(* Counting distance *)
IF bCount
    AND NOT fbFileHandler.bFileRead
THEN
	lrNoRetainDistance := lrNoRetainDistance + lrDistance;
	stRetainDistance.lrAllOverDistance := stCacheRetainDistance.lrAllOverDistance + lrNoRetainDistance;
	stRetainDistance.lrAfterResetDistance := stCacheRetainDistance.lrAfterResetDistance + lrNoRetainDistance;
END_IF


(* Write / read  file *)
fbFileHandler(
	bEnable := TRUE,
	dwDataBuffer := ADR(stRetainDistance),
	udnDataBufLen := SIZEOF(stRetainDistance),
	tTimeout := tTimeout,
	bError => bError,
	udnErrNo => udnErrNo
);

rtReset(
	CLK := NOT bSave AND bReset
);
IF rtReset.Q
THEN
	stRetainDistance.lrAfterResetDistance := 0;
	lrNoRetainDistance := 0;
END_IF

rtDeleteAll(
	CLK := NOT bSave AND bDeleteAll
);
IF rtDeleteAll.Q
THEN
	stRetainDistance.lrAllOverDistance := 0;
	stRetainDistance.lrAfterResetDistance := 0;
	stCacheRetainDistance.lrAllOverDistance := 0;
	stCacheRetainDistance.lrAfterResetDistance := 0;
	lrNoRetainDistance := 0;
END_IF

(* Counter distance mapping *)
lrAllOverDistance := stRetainDistance.lrAllOverDistance;
lrAfterResetDistance := stRetainDistance.lrAfterResetDistance;

END_FUNCTION_BLOCK

// ---- POUs/Tc2 Objects/Measurements/FB_TemperaturOK.TcPOU
FUNCTION_BLOCK FB_TemperaturOK
VAR_INPUT
	bEnable						:BOOL;			(* Enable FB signal *)
	bIn							:BOOL;			(* Temperature OK *)
	tTimeOutTempOK				:TIME := t#5s;		(* Temperature OK timeout *)
	tTimeOutTempNOK			:TIME := t#5s;		(* Temperature NOK timeout *)
END_VAR
VAR_OUTPUT
	bOut					:BOOL;			(* Temperature OK *)
	bError					:BOOL;			(* Error by temperature NOK *)
	udnErrorNo				:UDINT;
	udnMessageNo			:UDINT;
	sMsg					:STRING;
END_VAR
VAR
	bFirstTime			:BOOL;			(* First cycle *)
	tonDelayOK			:TON;			(* Temperatur delay ok *)
	tofWatchDog			:TOF;			(* Timer to off *)

END_VAR


IF NOT bFirstTime
THEN
	bError := FALSE;
	udnErrorNo := 0;
	udnMessageNo := 0;
	sMsg := '';
	tonDelayOK(
		IN := FALSE,
	          PT := tTimeOutTempOK
	);
	tofWatchDog(
		IN := FALSE,
	         PT := tTimeOutTempNOK
	);
	bFirstTime := TRUE;
END_IF;

(* Timer starts when came rising edge of signal *)
tonDelayOK(
	IN := bIn,
         PT := tTimeOutTempOK
);

tofWatchDog(
	IN := bIn,
         PT := tTimeOutTempNOK
);

IF tonDelayOK.Q
THEN
	bOut := TRUE;
    
ELSIF NOT tofWatchDog.Q
THEN
	bOut := FALSE;
    
END_IF;

END_FUNCTION_BLOCK

// ---- POUs/Tc2 Objects/Measurements/Oscat/T_PLC_MS.TcPOU
FUNCTION T_PLC_MS : DWORD
VAR CONSTANT
	debug			:BOOL := 0;
	N 				:INT := 0;
	offset 			:DWORD := 0;
END_VAR
VAR
	tx 				:TIME;
END_VAR

(*
version 1.2	16. nov 2008
programmer 	hugo
tested by	oscat

T_PLC_MS reads the internal PLC timer and return the time, it has the advantage to be able to set a debug mode 
and speed up the counter to test the plc timer overrun which occurs every 50 days respectively 25 days at siemens S7
this routine also allows to correct the behavior of s7 where the internal plc counter will not count all 32 bits.

*)

tx := TIME();
T_PLC_MS := TIME_TO_DWORD(Tx);
(* hier muss die korrektur für step7 stattfinden
plctime muss den vollen wertebereich von time ausnutzen:
wenn bei step7 time -24tage bis plus 24 tage ist dann muss der timer auch beim überlauf auf -24tage springen 
und auf keinen fall auf 0 !!!!
für siemens muss ein weiterer fb im main eingebunden werden der sicherstellt das alle 32 bits durchgezählt werden.
es kann nur ein fb sein den er muss sich das oberste (32te) bit merken.
oder etwa spring s7 bei überlauf auf -24 tage????? dann wäre keine korrektur nötig.
*)
IF debug
THEN
	T_PLC_MS := (SHL(T_PLC_MS,N) OR SHL(DWORD#1,N)-1) + OFFSET;
END_IF;

END_FUNCTION

// ---- POUs/Tc2 Objects/Safety/Fieldbus/FB_Fieldbus.TcPOU
FUNCTION_BLOCK FB_Fieldbus
(*

The function block used to control fieldbus.

Constructor: 		Patryk Panylo
Company:		E. Riexinger GmbH
Date:			23.04.2015
Version:			1.00

Date:			Revision:		Who:				Comment
dd.mm.yyyy		x.xx			Initials			comment

*)
VAR_INPUT
	(* Input variables / Eingang Variablen *)
	bEnable					:BOOL;						(* Enable FB signal *)
	unMasterState			:UINT;						(* Master state of fieldbus *)
														(* unFieldbus = 1 -> Sercos-Master:
															0xE001 = Phase 0
															0xE002 = Phase 1
															0xE003 = Phase 2
															0xE004 = Phase 3
															0xE005 = Phase 4
															0xE008 = Break
															0xE011 = Phase switch 0 -> 1
															0xE012 = Phase switch 1 -> 2
															0xE013 = Phase switch 2 -> 3
															0xE014 = Phase switch 3 -> 4
					
														  uiFieldbus = 2 -> EtherCat Master:
															0x0001 = Link error
															0x0002 = I/O locked after link error (I/O reset required)
															0x0004 = Link error (redundancy adapter)
															0x0008 = Missing one frame (redundancy mode)
															0x0010 = Out of send resources (I/O reset required)
															0x0020 = Watchdog triggered
															0x0040 = Ethernet driver (miniport) not found
															0x0080 = I/O reset active
															0x0100 = At least one device in 'INIT' state
															0x0200 = At least one device in 'PRE-OP' state
															0x0400 = At least one device in 'SAFE-OP' state
															0x0800 = At least one device indicates an error state
															0x1000 = DC not in sync
														*)
	unSlaveState				:ARRAY[1..unSlaveNo] OF UINT;	(* State of slaves periphery / Status des Periphery
														uiFieldbus = 2 -> EtherCat Master:
															0x___1 = Slave in 'INIT' state
															0x___2 = Slave in 'PREOP' state
															0x___3 = Slave in 'BOOT' state
															0x___4 = Slave in 'SAFEOP' state
															0x___8 = Slave in 'OP' state
															0x001_ = Slave signals error
															0x002_ = Invalid vendorId, productCode... read
															0x004_ = Initialization error occurred
															0x008_ = Slave disabled
															0x010_ = Slave not present
															0x020_ = Slave signals link error
															0x040_ = Slave signals missing link
															0x080_ = Slave signals unexpected link
															0x100_ = Communication port A
															0x200_ = Communication port B
															0x400_ = Communication port C
															0x800_ = Communication port D
													*)
	tAdsTimeOut				:TIME := t#5s;				(* Timeout for ADS commando *)
END_VAR
VAR_OUTPUT
	(* Output variables / Ausgang Variablen *)
	sDeviceNetId				:T_AmsNetId ;			(* Fieldbus master ams net id*)
	bInitReady				:BOOL;					(* Fieldbus master initialisation is complete*)
	bBreak					:BOOL;					(* Fieldbus break *)
	bError					:BOOL;					(* Error by no air pressure *)
	udnErrorNo				:UDINT;
	udnMessageNo			:UDINT;
	sMsg					:STRING;
END_VAR
VAR
	(* Enummerations *)

	(* Variables *)
	unSlaveCounter			:UINT;					(* Slave counter *)
	bBreakMasterState		:BOOL;					(* Fieldbus master break *)
	bBreakSlaveState			:BOOL;					(* Fieldbus slave break *)

	(* References *)

	(* Interfaces *)

	(* Instances *)
	fbGetDeviceNetId			:IOF_GetDeviceNetId; 		(* Get the device net id from the device ID *)
	fbGetDeviceType			:IOF_GetDeviceType; 		(* Get the device type from the device ID *)
END_VAR
VAR CONSTANT
	unSlaveNo				:UINT := 32;				(* Number of slaves in Fieldbus *)
END_VAR

IF NOT bEnable
THEN
	fbGetDeviceNetId(START := FALSE);
	fbGetDeviceType(START := FALSE);
	bInitReady := FALSE;
	bBreak := FALSE;
	bError := FALSE;
	udnErrorNo := 0;
	udnMessageNo := 0;
	sMsg := '';
	RETURN;
END_IF;

(* Get the device net id from the device ID *)
fbGetDeviceNetId(
	NETID := '',
	DEVICEID := 1,
	START := TRUE,
	TMOUT := tAdsTimeOut
);

(* Get the device type from the device ID *)
fbGetDeviceType(
	NETID := '',
	DEVICEID := 1,
	START := TRUE,
	TMOUT := tAdsTimeOut
);

(* Get the device net id from the device ID *)
IF NOT fbGetDeviceNetId.BUSY 											(* No error *)
     AND NOT fbGetDeviceNetId.ERR
THEN
	sDeviceNetId := fbGetDeviceNetId.DeviceNetId;							(* Device net id *)

	(* Get the device type from the device ID *)
	IF NOT fbGetDeviceType.BUSY 										(* No error *)
	     AND NOT fbGetDeviceType.ERR
	THEN

		CASE fbGetDeviceType.IODeviceType
		OF
			48: (* IODEVICETYPE_FC7500 	:= 48,  Beckhoff-SERCOS-PCI *)
				bError := FALSE;
				udnErrorNo := 0;											(* Error number *)
				bInitReady := unMasterState = 16#E005; 						(* Actual Phase is 4 *)
				bBreak := unMasterState = 16#E008;							(* Interrupt / Broke *)
			94: (* IODEVICETYPE_EtherCAT := 94,  Beckhoff-EtherCAT-PCI *)
				bError := FALSE;
				udnErrorNo := 0;											(* Error number *)
				bInitReady := unMasterState = 16#0000; 						(* Actual master state is OP *)

				bBreakMasterState :=  unMasterState <> 16#0000;				(* Fieldbus master break *)

				IF bInitReady
				THEN
					bBreakSlaveState := FALSE;							(* Fieldbus slave break *)

					FOR unSlaveCounter :=1 TO unSlaveNo
					DO
						bBreakSlaveState := unSlaveState[unSlaveCounter] <> 16#0000
										     AND unSlaveState[unSlaveCounter] <> 16#0008;

						IF bBreakSlaveState
						THEN
							EXIT;
						END_IF

					END_FOR;
				END_IF

				bBreak := bBreakMasterState 								(* Interrupt / Broke *)
						 OR bBreakSlaveState;

		ELSE (* IDLE *)
			bInitReady := FALSE;
			bBreak := FALSE;
			bError := TRUE;
			udnErrorNo := 1;																			(* Error number *)
			sMsg := CONCAT('Unidentified fieldbus:', DINT_TO_STRING(fbGetDeviceType.IODeviceType));		(* Description error *)
		END_CASE;

	ELSIF NOT fbGetDeviceType.BUSY
		   AND fbGetDeviceType.ERR
	THEN
		bError := TRUE;
		udnErrorNo := 2;																				(* Error number *)
		sMsg := CONCAT('Fehler beim Lesen über ADS: ', UDINT_TO_STRING(fbGetDeviceType.ERRID));		(* Description error *)
		fbGetDeviceType(START := FALSE);
	END_IF;

ELSIF NOT fbGetDeviceNetId.BUSY
	    AND fbGetDeviceNetId.ERR
THEN
	bError := TRUE;
	udnErrorNo := 3;																					(* Error number *)
	sMsg := CONCAT('Fehler beim Lesen über ADS: ', UDINT_TO_STRING(fbGetDeviceNetId.ERRID));			(* Description error *)
	fbGetDeviceNetId(START := FALSE);
END_IF;

END_FUNCTION_BLOCK

// ---- POUs/Tc2 Objects/Signals/Force Input/FB_ForceBit.TcPOU
FUNCTION_BLOCK FB_ForceBit
(*

Forcing the input bit through pointer.
IO variables in VAR_CONFIG are generated automatically by TwinCAT - read only
Matching variable must be with  %I* declarated.

Constructor: 		Patryk Panylo
Company:		E. Riexinger GmbH
Date:			28.10.2013
Version:			1.00

Date:			Revision:		Who:				Comment
dd.mm.yyyy		x.xx			Initials			comment

*)
VAR_INPUT
	bEnable						:BOOL; 							(* Enable FB *)
	dwBitAddr					:DWORD;						(* The address of input argument in a DWORD: BITADR(Input) where e.g Input = %IX0.1 *)
	bForceInState				:BOOL;							(* Force input state *)
	tDelayOn					:TIME;							(* Delay signal on *)
	tDelayOff						:TIME;							(* Delay signal off *)
END_VAR
VAR_OUTPUT
END_VAR
VAR
	pByteAddr					:POINTER TO BYTE;
	byCurrentInState				:BYTE;							(* Current input state *)
	byBitMask					:BYTE;

	tonDelayOn					:TON;
	tonDelayOff					:TOF;

END_VAR

IF NOT bEnable
THEN
	RETURN;
END_IF

(* Delay on signal *)
tonDelayOn(
	IN := bForceInState,
	PT := tDelayOn
);

(* Delay off signal *)
tonDelayOff(
	IN := tonDelayOn.Q,
	PT := tDelayOff
);

pByteAddr := ADR(%IB0) + (dwBitAddr / 8);
byCurrentInState := pByteAddr^;

byBitMask := SHL(BYTE#1, (dwBitAddr AND 2#00000111));

IF tonDelayOff.Q
THEN
	pByteAddr^ := byCurrentInState OR byBitMask;
ELSE
	pByteAddr^ := byCurrentInState AND NOT byBitMask;
END_IF

END_FUNCTION_BLOCK

// ---- POUs/Tc2 Objects/Signals/Force Input/FB_ForceByte.TcPOU
FUNCTION_BLOCK FB_ForceByte
(*

Forcing the input bit through pointer.
IO variables in VAR_CONFIG are generated automatically by TwinCAT - read only
Matching variable must be with  %I* declarated.

Constructor: 		Patryk Panylo
Company:		E. Riexinger GmbH
Date:			28.10.2013
Version:			1.00

Date:			Revision:		Who:				Comment
dd.mm.yyyy		x.xx			Initials			comment

*)
VAR_INPUT
	bEnable						:BOOL; 							(* Enable FB *)
	dwAddr						:DWORD;						(* The address of input argument in a DWORD: ADR(Input) where e.g Input = %IB *)
	bForceInState				:BOOL;							(* Force input state *)
	tDelayOn					:TIME;							(* Delay signal on *)
	tDelayOff						:TIME;							(* Delay signal off *)
END_VAR
VAR_OUTPUT
END_VAR
VAR
	pByteAddr					:POINTER TO BYTE;
	byCurrentInState				:BYTE;							(* Current input state *)
	byBitMask					:BYTE;

	tonDelayOn					:TON;
	tonDelayOff					:TOF;

END_VAR

IF NOT bEnable
THEN
	RETURN;
END_IF

(* Delay on signal *)
tonDelayOn(
	IN := bForceInState,
	PT := tDelayOn
);

(* Delay off signal *)
tonDelayOff(
	IN := tonDelayOn.Q,
	PT := tDelayOff
);

pByteAddr := dwAddr;
byCurrentInState := pByteAddr^;

byBitMask := 2#00000001;

IF tonDelayOff.Q
THEN
	pByteAddr^ := byCurrentInState OR byBitMask;
ELSE
	pByteAddr^ := byCurrentInState AND NOT byBitMask;
END_IF

END_FUNCTION_BLOCK

// ---- POUs/Tc2 Objects/Signals/Handling/F_SignalHandling.TcPOU
FUNCTION F_SignalHandling : BOOL
VAR_INPUT
	(* Input variables / Eingang Variablen *)
	bEnable					:BOOL;						(* Enable FB signal *)
	bIn						:BOOL;						(* Input signal *)
END_VAR
VAR
END_VAR

IF NOT bEnable
THEN
	F_SignalHandling := FALSE;
    	RETURN;
END_IF;

F_SignalHandling := bIn;                     (* Set output *)

END_FUNCTION

// ---- POUs/Tc2 Objects/Signals/Ramp Generators/FB_RampDirector.TcPOU
FUNCTION_BLOCK FB_RampDirector
(*

Frequency division

Constructor: 		Patryk Panylo
Company:		E. Riexinger GmbH
Date:			14.11.2012
Version:			1.00

Date:			Revision:		Who:				Comment
dd.mm.yyyy		x.xx			Initials			comment

*)

VAR_INPUT
	bEnable						:BOOL;						(* Function block enable *)
	bExecute					:BOOL;						(* Execut the function block *)
	bDirection					:BOOL;						(* Rising = 1, Falling = 0 *)
	bSet						:BOOL;						(* Set output to 65535 *)
	bReset						:BOOL;						(* Reset output to 0 *)
	tRiseTime					:TIME;						(* Rise time of ramp *)
	tFallTime					:TIME;						(* Fall time of ramp *)
	rHighLimit					:REAL;						(* High limit of ramp *)
	rLowLimit						:REAL;						(* Low limit of ramp *)
	rNoLimit						:REAL;						(* No limit value active if rise and fall time no active *)
END_VAR
VAR_OUTPUT
	wRVOut						:WORD;						(* Ramp value, 100% = 65535 *)
	rPVOut						:REAL;						(* Judgment Value *)
	nPVOut						:INT;						(* Judgment Value *)
	bLowLevel					:BOOL;						(* Low level reached *)
	bHighLevel					:BOOL;						(* High level reached *)
	bDone						:BOOL;						(* Program done *)
	bBusy 						:BOOL;						(* Program busy *)
	bError 						:BOOL;						(* Program error *)
END_VAR
VAR
	fbRampGen					:FB_RMP_W;					(* Ramp generator *)

	rCacheLowLimit				:REAL;
	rCacheHighLimit				:REAL;

	rtExecute						:R_TRIG;
	etRampGenerator				:ET_RampGenerator;
END_VAR


IF NOT bEnable
THEN
	bDone := FALSE;                                     (* Program done *)
	bBusy := FALSE;                                     (* Program not busy *)
	bError := FALSE;                                    (* Program not error *)
	
	rtExecute(CLK := FALSE);

	fbRampGen(
		bEnable := FALSE,
		bReset := bReset,
		bSet := bSet,
		wRVOut => wRVOut
	);

	RETURN;
END_IF;

rtExecute(CLK := bExecute);

IF rtExecute.Q
THEN
	fbRampGen(
		bEnable := FALSE,
		bDirection := bDirection,
		bSet := FALSE,
		bReset := FALSE,
		tRampTime := T#0ms
	);
	
	etRampGenerator := ET_RampGenerator_eWaitExecute;						(* Next step *)

END_IF

(* Reset ramp *)
IF (tFallTime = t#0s
    AND tRiseTime <> t#0s
    AND bExecute
    AND NOT bDirection)
    OR bReset
THEN
	fbRampGen.bReset := TRUE;
	wRVOut := fbRampGen.wRVOut;
ELSE
	fbRampGen.bReset := FALSE;
END_IF;

(* Set ramp *)
IF (tRiseTime = t#0s
    AND tFallTime <> t#0s
    AND bExecute
    AND bDirection)
    OR bSet
THEN
	fbRampGen.bSet := TRUE;
ELSE
	fbRampGen.bSet := FALSE;
END_IF;

(* Call ramp generator *)
fbRampGen(
	bDirection := bDirection,
	tRampTime := SEL(bDirection, tFallTime, tRiseTime),
	bLowLevel => bLowLevel,
	bHighLevel => bHighLevel
);

IF fbRampGen.bReset
    OR fbRampGen.bSet
THEN
	wRVOut := fbRampGen.wRVOut;
END_IF;

CASE etRampGenerator OF
        
	ET_RampGenerator_eWaitExecute:
		bDone := FALSE;                                     (* Program done *)
		bBusy := FALSE;                                     (* Program not  busy *)
		bError := FALSE;                                    (* Program not error *)

		fbRampGen.bEnable := FALSE;
		
		IF rtExecute.Q
		THEN
			bDone := FALSE;                                     (* Program done *)
			bBusy := TRUE;                                 	 	(* Program not busy *)

			IF tRiseTime = t#0s
    			     AND tFallTime = t#0s
			THEN
				fbRampGen.bEnable := FALSE;

				rCacheLowLimit := rNoLimit;
				rCacheHighLimit := rNoLimit;

				etRampGenerator := ET_RampGenerator_eDone;         (* Next step *)
			ELSE
				fbRampGen.bEnable := TRUE;

				rCacheLowLimit := rLowLimit;
				rCacheHighLimit := rHighLimit;

				etRampGenerator := ET_RampGenerator_eRunning;           (* Next step *)
			END_IF
		END_IF

	ET_RampGenerator_eRunning:
		IF fbRampGen.bBusy
		THEN
			wRVOut := fbRampGen.wRVOut;
		
			etRampGenerator := ET_RampGenerator_eWaiting;           (* Next step *)
		END_IF
        
	ET_RampGenerator_eWaiting:
		IF fbRampGen.bBusy
		THEN
			wRVOut := fbRampGen.wRVOut;
		ELSE
			fbRampGen.bEnable := FALSE;
		
			etRampGenerator := ET_RampGenerator_eDone;         (* Next step *)
		END_IF		

	ET_RampGenerator_eDone:
		bDone := TRUE;                                      (* Program done *)
		bBusy := FALSE;                                     (* Program not busy *)
		
		etRampGenerator := ET_RampGenerator_eNotExecute;            (* Next step *)
        
	ET_RampGenerator_eError:
		bDone := FALSE;                                     (* Program done *)
		bBusy := FALSE;                                     (* Program not busy *)
		bError := TRUE;                                     (* Program error *)
		
		etRampGenerator := ET_RampGenerator_eNotExecute;            (* Next step *)
        
	ET_RampGenerator_eNotExecute:
	IF NOT bExecute
	THEN
		bDone := FALSE;                                     (* Program done *)
		bBusy := FALSE;                                     (* Program not busy *)
		bError := FALSE;                                    (* Program not error *)

		wRVOut := fbRampGen.wRVOut;
	
		etRampGenerator := ET_RampGenerator_eWaitExecute;               (* Next step *)

	END_IF;
END_CASE;

rPVOut := F_WordToRange(
			wWord := wRVOut,
			rLowLimit := rCacheLowLimit,
			rHighLimit := rCacheHighLimit
		);

nPVOut := REAL_TO_INT(rPVOut);

END_FUNCTION_BLOCK

// ---- POUs/Tc2 Objects/Signals/Watchdog/FB_SignalWatchdog2.TcPOU
FUNCTION_BLOCK FB_SignalWatchdog2
VAR_INPUT
	bEnable					:BOOL;			(* Enable FB signal *)
	bIn						:BOOL;			(* Input *)
	tTimeOutHigh				:TIME := t#5s;		(* Input high timeout *)
	tTimeOutLow				:TIME := t#5s;		(* Input low timeout *)
END_VAR
VAR_OUTPUT
	bOut					:BOOL;			(* Output *)
	bError					:BOOL;			(* Error *)
	udnErrorNo				:UDINT;
	udnMessageNo			:UDINT;
	sMsg					:STRING;
END_VAR
VAR
	bFirstTime				:BOOL;			(* First cycle *)
	tonDelay					:TON;			(* Delay *)
	tofWatchDog				:TOF;			(* Timer to off *)

END_VAR


IF NOT bFirstTime
THEN
	bError := FALSE;
	udnErrorNo := 0;
	udnMessageNo := 0;
	sMsg := '';
	tonDelay(
		IN := FALSE,
	          PT := tTimeOutHigh
	);
	tofWatchDog(
		IN := FALSE,
	         PT := tTimeOutLow
	);
	bFirstTime := TRUE;
END_IF;

(* Timer starts when came rising edge of signal *)
tonDelay(
	IN := bIn,
         PT := tTimeOutHigh
);

tofWatchDog(
	IN := bIn,
         PT := tTimeOutLow
);

IF tonDelay.Q
THEN
	bOut := TRUE;
    
ELSIF NOT tofWatchDog.Q
THEN
	bOut := FALSE;
    
END_IF;

END_FUNCTION_BLOCK

// ---- POUs/Tc2 Objects/String/F_RealToStrf.TcPOU
FUNCTION F_RealToStrf : STRING(20)
VAR_INPUT
	IN : REAL;
	N : INT;
	D : STRING(1);
END_VAR
VAR
	O: REAL;
	i: INT;
END_VAR

(*
version 1.8	2. jan 2012
programmer 	hugo
tested by	oscat

Real_to_strf converts a Real to a fixed length String.
the string will be filles with zeroes to achieve the fixed length N after the decimal separator.
the input parameter specifies the decimal separator to be used in the output string.

*)

(* LIMIT N to 0 .. 7 *)
N := LIMIT(0,N,7);
(* round the input to N digits and convert to string *)
O := ABS(in) * F_Exp10(N);
F_RealToStrf := DINT_TO_STRING(REAL_TO_DINT(O));
(* add zeroes in front to make sure sting is at least 8 digits long *)
FOR i := LEN(F_RealToStrf) TO N DO F_RealToStrf := CONCAT('0', F_RealToStrf); END_FOR;
(* add a dot if n > 0 *)
IF n > 0 THEN F_RealToStrf := INSERT(F_RealToStrf, D, LEN(F_RealToStrf) - N); END_IF;
(* add a minus sign if in is negative *)
IF in < 0 THEN F_RealToStrf := CONCAT('-', F_RealToStrf); END_IF;

END_FUNCTION

// ---- POUs/Tc3 Objects/Alarm/FB_Alarm_1.TcPOU
FUNCTION_BLOCK FB_Alarm_1
VAR_INPUT
	(* Input variables / Eingang Variablen *)
	bEnable					:BOOL;						(* Enable FB signal *)
	bNoEStop				:BOOL;						(* Emergency stop *)
	bReset					:BOOL;						(* Reset *)
	dtDateTime 				:DATE_AND_TIME;				(* Actual date and time *)
	nFatalErrorMaxIdx		:INT;						(* Maximal index of  using alarms *)
	nErrorMaxIdx			:INT;						(* Maximal index of  using alarms *)
	nWarningMaxIdx			:INT;						(* Maximal index of  using alarms *)
	nMessageMaxIdx			:INT;						(* Maximal index of  using alarms *)
	nHintMaxIdx				:INT;						(* Maximal index of  using alarms *)
	stAlarmIn				:ST_AlarmIn;					(* Alarm input *)
END_VAR
VAR_OUTPUT
	(* Output variables / Ausgang Variablen *)
END_VAR
VAR_IN_OUT
	(* Input Output variables / Ausgang Variablen *)
	stAlarmOut				:ST_AlarmOut;				(* Alarm output *)
END_VAR
VAR
	(* Enummerations *)

	(* Variables *)
	arfbFatalError				:ARRAY[0..nALARM_MAX_NO] OF FB_FatalError;
	arfbError					:ARRAY[0..nALARM_MAX_NO] OF FB_Error;
	arfbWarning					:ARRAY[0..nALARM_MAX_NO] OF FB_Warning;
	arfbMessage					:ARRAY[0..nALARM_MAX_NO] OF FB_Message;
	arfbHint					:ARRAY[0..nALARM_MAX_NO] OF FB_Hint;

	nInc						:INT;

	(* References *)

	(* Interfaces *)

	(* Instances *)
	rtNoEStop				:R_TRIG;
	tonNoEStopDelay			:TON;
END_VAR

IF NOT bEnable
THEN
    RETURN;
END_IF;

IF dtDateTime = DT#1970-01-01-00:00
THEN
	RETURN;
END_IF

tonNoEStopDelay(
	IN := bNoEStop, 
	PT := T#1S
);
rtNoEStop(CLK := tonNoEStopDelay.Q);

stAlarmOut.bFatalError := FALSE;
stAlarmOut.bError := FALSE;
stAlarmOut.bWarning := FALSE;
stAlarmOut.bMessage := FALSE;
stAlarmOut.bHint := FALSE;

IF nFatalErrorMaxIdx > nALARM_MAX_NO
THEN
	nFatalErrorMaxIdx := nALARM_MAX_NO;
END_IF
FOR nInc := 0 TO nFatalErrorMaxIdx
DO
	(* ************************ FatalError ************************ *)
	stAlarmIn.arbFatalError[nInc].enType := ET_AlarmType.eFatalError;
	stAlarmIn.arbFatalError[nInc].dtDateTime := dtDateTime;
	
	arfbFatalError[nInc](
		bEnable := TRUE,
		stAlarmIn := stAlarmIn.arbFatalError[nInc]
	);

	stAlarmOut.arbFatalError[nInc].bActive := arfbFatalError[nInc].stAlarmOut.bActive;
	stAlarmOut.arbFatalError[nInc].dtDateTime := arfbFatalError[nInc].stAlarmOut.dtDateTime;
	stAlarmOut.arbFatalError[nInc].enType := arfbFatalError[nInc].stAlarmOut.enType;
	stAlarmOut.arbFatalError[nInc].dnCode := arfbFatalError[nInc].stAlarmOut.dnCode;
	
	stAlarmOut.bFatalError := stAlarmOut.bFatalError OR (stAlarmOut.arbFatalError[nInc].bActive > 0);
END_FOR

IF nErrorMaxIdx > nALARM_MAX_NO
THEN
	nErrorMaxIdx := nALARM_MAX_NO;
END_IF
FOR nInc := 0 TO nErrorMaxIdx
DO
	(* ************************ Error ************************ *)
	stAlarmIn.arbError[nInc].enType := ET_AlarmType.eError;
	stAlarmIn.arbError[nInc].dtDateTime := dtDateTime;
	
	arfbError[nInc](
		bEnable := TRUE,
		bReset := bReset OR rtNoEStop.Q,
		stAlarmIn := stAlarmIn.arbError[nInc]
	);

	stAlarmOut.arbError[nInc].bActive := arfbError[nInc].stAlarmOut.bActive;
	stAlarmOut.arbError[nInc].dtDateTime := arfbError[nInc].stAlarmOut.dtDateTime;
	stAlarmOut.arbError[nInc].enType := arfbError[nInc].stAlarmOut.enType;
	stAlarmOut.arbError[nInc].dnCode := arfbError[nInc].stAlarmOut.dnCode;
	
	stAlarmOut.bError := stAlarmOut.bError OR (stAlarmOut.arbError[nInc].bActive > 0);
END_FOR

IF nWarningMaxIdx > nALARM_MAX_NO
THEN
	nWarningMaxIdx := nALARM_MAX_NO;
END_IF
FOR nInc := 0 TO nWarningMaxIdx
DO
	(* ************************ Warning ************************ *)
	stAlarmIn.arbWarning[nInc].enType := ET_AlarmType.eWarning;
	stAlarmIn.arbWarning[nInc].dtDateTime := dtDateTime;
	
	arfbWarning[nInc](
		bEnable := TRUE,
		bReset := bReset OR rtNoEStop.Q,
		stAlarmIn := stAlarmIn.arbWarning[nInc]
	);
	
	stAlarmOut.arbWarning[nInc].bActive := arfbWarning[nInc].stAlarmOut.bActive;
	stAlarmOut.arbWarning[nInc].dtDateTime := arfbWarning[nInc].stAlarmOut.dtDateTime;
	stAlarmOut.arbWarning[nInc].enType := arfbWarning[nInc].stAlarmOut.enType;
	stAlarmOut.arbWarning[nInc].dnCode := arfbWarning[nInc].stAlarmOut.dnCode;
	
	stAlarmOut.bWarning := stAlarmOut.bWarning OR (stAlarmOut.arbWarning[nInc].bActive > 0);
END_FOR

IF nMessageMaxIdx > nALARM_MAX_NO
THEN
	nMessageMaxIdx := nALARM_MAX_NO;
END_IF
FOR nInc := 0 TO nMessageMaxIdx
DO
	(* ************************ Message ************************ *)
	stAlarmIn.arbMessage[nInc].enType := ET_AlarmType.eMessage;
	stAlarmIn.arbMessage[nInc].dtDateTime := dtDateTime;
	
	arfbMessage[nInc](
		bEnable := TRUE,
		stAlarmIn := stAlarmIn.arbMessage[nInc]
	);
	
	stAlarmOut.arbMessage[nInc].bActive := arfbMessage[nInc].stAlarmOut.bActive;
	stAlarmOut.arbMessage[nInc].dtDateTime := arfbMessage[nInc].stAlarmOut.dtDateTime;
	stAlarmOut.arbMessage[nInc].enType := arfbMessage[nInc].stAlarmOut.enType;
	stAlarmOut.arbMessage[nInc].dnCode := arfbMessage[nInc].stAlarmOut.dnCode;
		
	stAlarmOut.bMessage := stAlarmOut.bMessage OR (stAlarmOut.arbMessage[nInc].bActive > 0);
END_FOR

IF nHintMaxIdx > nALARM_MAX_NO
THEN
	nHintMaxIdx := nALARM_MAX_NO;
END_IF
FOR nInc := 0 TO nHintMaxIdx
DO
	(* ************************ Hint ************************ *)
	stAlarmIn.arbMessage[nInc].enType := ET_AlarmType.eMessage;
	stAlarmIn.arbMessage[nInc].dtDateTime := dtDateTime;
	
	arfbHint[nInc](
		bEnable := TRUE,
		stAlarmIn := stAlarmIn.arbHint[nInc]
	);

	stAlarmOut.arbHint[nInc].bActive := arfbHint[nInc].stAlarmOut.bActive;
	stAlarmOut.arbHint[nInc].dtDateTime := arfbHint[nInc].stAlarmOut.dtDateTime;
	stAlarmOut.arbHint[nInc].enType := arfbHint[nInc].stAlarmOut.enType;
	stAlarmOut.arbHint[nInc].dnCode := arfbHint[nInc].stAlarmOut.dnCode;
	
	stAlarmOut.bHint := stAlarmOut.bHint OR (stAlarmOut.arbHint[nInc].bActive > 0);
END_FOR

END_FUNCTION_BLOCK

// ---- POUs/Tc3 Objects/Alarm/FB_Error_1.TcPOU
FUNCTION_BLOCK FB_Error_1
VAR_INPUT
	(* Input variables / Eingang Variablen *)
	bEnable					:BOOL;						(* Enable FB signal *)
	bReset					:BOOL;						(* Reset *)
	stAlarmIn				:ST_AlarmProperties;				(* Alarm output *)
END_VAR
VAR_OUTPUT
	(* Output variables / Ausgang Variablen *)
	stAlarmOut				:ST_AlarmProperties;				(* Alarm output *)
END_VAR
VAR_IN_OUT

END_VAR
VAR
	(* Enummerations *)

	(* Variables *)

	(* References *)

	(* Interfaces *)

	(* Instances *)

END_VAR

(* Check method enabled *)
IF NOT bEnable
THEN
	RETURN;
END_IF;

IF bReset
THEN
	IF stAlarmOut.bActive
	THEN
		stAlarmOut.bActive := FALSE;
		//stAlarmOut.enType := ET_AlarmType.eIdle;
		//stAlarmOut.dtDateTime := DT#1970-01-01-00:00;
		//stAlarmOut.dnCode := 0;
	END_IF;
ELSE
	IF stAlarmIn.bActive
	    AND NOT stAlarmOut.bActive
	THEN
		stAlarmOut.bActive := TRUE;
		stAlarmOut.enType := stAlarmIn.enType;
		stAlarmOut.dtDateTime := stAlarmIn.dtDateTime;
		stAlarmOut.dnCode := stAlarmIn.dnCode;
	END_IF;
END_IF;

END_FUNCTION_BLOCK

// ---- POUs/Tc3 Objects/Alarm/FB_FatalError_1.TcPOU
FUNCTION_BLOCK FB_FatalError_1
VAR_INPUT
	(* Input variables / Eingang Variablen *)
	bEnable					:BOOL;						(* Enable FB signal *)
	stAlarmIn				:ST_AlarmProperties;				(* Alarm output *)
END_VAR
VAR_OUTPUT
	(* Output variables / Ausgang Variablen *)
	stAlarmOut				:ST_AlarmProperties;				(* Alarm output *)
END_VAR
VAR_IN_OUT

END_VAR
VAR
	(* Enummerations *)

	(* Variables *)

	(* References *)

	(* Interfaces *)

	(* Instances *)
	rtAlarm					:R_TRIG;
	ftAlarm					:F_TRIG;
END_VAR

(* Check method enabled *)
IF NOT bEnable
THEN
	RETURN;
END_IF;

rtAlarm(CLK := stAlarmIn.bActive);
ftAlarm(CLK := stAlarmIn.bActive);

IF rtAlarm.Q
THEN
	stAlarmOut.bActive := TRUE;
	stAlarmOut.enType := stAlarmIn.enType;
	stAlarmOut.dtDateTime := stAlarmIn.dtDateTime;
	stAlarmOut.dnCode := stAlarmIn.dnCode;
	
ELSIF ftAlarm.Q
THEN
	stAlarmOut.bActive := FALSE;
	//stAlarmOut.enType := ET_AlarmType.eIdle;
	//stAlarmOut.dtDateTime := DT#1970-01-01-00:00;
	//stAlarmOut.dnCode := 0;
END_IF;

END_FUNCTION_BLOCK

// ---- POUs/Tc3 Objects/Alarm/FB_Hint_1.TcPOU
FUNCTION_BLOCK FB_Hint_1
VAR_INPUT
	(* Input variables / Eingang Variablen *)
	bEnable					:BOOL;						(* Enable FB signal *)
	stAlarmIn				:ST_AlarmProperties;				(* Alarm output *)
END_VAR
VAR_OUTPUT
	(* Output variables / Ausgang Variablen *)
	stAlarmOut				:ST_AlarmProperties;				(* Alarm output *)
END_VAR
VAR_IN_OUT

END_VAR
VAR
	(* Enummerations *)

	(* Variables *)

	(* References *)

	(* Interfaces *)

	(* Instances *)
	rtAlarm					:R_TRIG;
	ftAlarm					:F_TRIG;
END_VAR

(* Check method enabled *)
IF NOT bEnable
THEN
	RETURN;
END_IF;

rtAlarm(CLK := stAlarmIn.bActive);
ftAlarm(CLK := stAlarmIn.bActive);

IF rtAlarm.Q
THEN
	stAlarmOut.bActive := TRUE;
	stAlarmOut.enType := stAlarmIn.enType;
	stAlarmOut.dtDateTime := stAlarmIn.dtDateTime;
	stAlarmOut.dnCode := stAlarmIn.dnCode;
    
ELSIF ftAlarm.Q
THEN
	stAlarmOut.bActive := FALSE;
	//stAlarmOut.enType := ET_AlarmType.eIdle;
	//stAlarmOut.dtDateTime := DT#1970-01-01-00:00;
	//stAlarmOut.dnCode := 0;	
END_IF;

END_FUNCTION_BLOCK

// ---- POUs/Tc3 Objects/Alarm/FB_Message_1.TcPOU
FUNCTION_BLOCK FB_Message_1
VAR_INPUT
	(* Input variables / Eingang Variablen *)
	bEnable					:BOOL;						(* Enable FB signal *)
	stAlarmIn				:ST_AlarmProperties;				(* Alarm output *)
END_VAR
VAR_OUTPUT
	(* Output variables / Ausgang Variablen *)
	stAlarmOut				:ST_AlarmProperties;				(* Alarm output *)
END_VAR
VAR_IN_OUT

END_VAR
VAR
	(* Enummerations *)

	(* Variables *)

	(* References *)

	(* Interfaces *)

	(* Instances *)
	rtAlarm					:R_TRIG;
	ftAlarm					:F_TRIG;
END_VAR

(* Check method enabled *)
IF NOT bEnable
THEN
	RETURN;
END_IF;

rtAlarm(CLK := stAlarmIn.bActive);
ftAlarm(CLK := stAlarmIn.bActive);

IF rtAlarm.Q
THEN
	stAlarmOut.bActive := TRUE;
	stAlarmOut.enType := stAlarmIn.enType;
	stAlarmOut.dtDateTime := stAlarmIn.dtDateTime;
	stAlarmOut.dnCode := stAlarmIn.dnCode;
    
ELSIF ftAlarm.Q
THEN
	stAlarmOut.bActive := FALSE;
	//stAlarmOut.enType := ET_AlarmType.eIdle;
	//stAlarmOut.dtDateTime := DT#1970-01-01-00:00;
	//stAlarmOut.dnCode := 0;
END_IF;

END_FUNCTION_BLOCK

// ---- POUs/Tc3 Objects/Alarm/FB_Warning_1.TcPOU
FUNCTION_BLOCK FB_Warning_1
VAR_INPUT
	(* Input variables / Eingang Variablen *)
	bEnable					:BOOL;						(* Enable FB signal *)
	bReset					:BOOL;						(* Reset *)
	stAlarmIn				:ST_AlarmProperties;				(* Alarm output *)
END_VAR
VAR_OUTPUT
	(* Output variables / Ausgang Variablen *)
	stAlarmOut				:ST_AlarmProperties;				(* Alarm output *)
END_VAR
VAR_IN_OUT

END_VAR
VAR
	(* Enummerations *)

	(* Variables *)

	(* References *)

	(* Interfaces *)

	(* Instances *)

END_VAR

(* Check method enabled *)
IF NOT bEnable
THEN
	RETURN;
END_IF;

IF bReset
THEN
	IF stAlarmOut.bActive
	THEN
		stAlarmOut.bActive := FALSE;
		//stAlarmOut.enType := ET_AlarmType.eIdle;
		//stAlarmOut.dtDateTime := DT#1970-01-01-00:00;
		//stAlarmOut.dnCode := 0;
	END_IF;
	
ELSE
	IF stAlarmIn.bActive
	    AND NOT stAlarmOut.bActive
	THEN
		stAlarmOut.bActive := TRUE;
		stAlarmOut.enType := stAlarmIn.enType;
		stAlarmOut.dtDateTime := stAlarmIn.dtDateTime;
		stAlarmOut.dnCode := stAlarmIn.dnCode;
	END_IF;
	
END_IF;

END_FUNCTION_BLOCK

// ---- POUs/Tc3 Objects/Automation/Axis/F_ChkAllAxisCoupled_1.TcPOU
FUNCTION F_ChkAllAxisCoupled_1 : BOOL
(*

The function used to detect if all axis are coupled.

Constructor: 		Patryk Panylo
Company:		E. Riexinger GmbH
Date:			23.04.2015
Version:			1.00

Date:			Revision:		Who:				Comment
dd.mm.yyyy		x.xx			Initials			comment

*)
VAR_INPUT
	(* Input variables / Eingang Variablen *)
	bEnable						:BOOL;					(* Signal FB enable *)
	bAxis1Coupled				:BOOL;					(* Axis coupled *)
	bAxis2Coupled				:BOOL;					(* Axis coupled *)
	bAxis3Coupled				:BOOL;					(* Axis coupled *)
	bAxis4Coupled				:BOOL;					(* Axis coupled *)
	bAxis5Coupled				:BOOL;					(* Axis coupled *)
	bAxis6Coupled				:BOOL;					(* Axis coupled *)
	bAxis7Coupled				:BOOL;					(* Axis coupled *)
	bAxis8Coupled				:BOOL;					(* Axis coupled *)
	bAxis9Coupled				:BOOL;					(* Axis coupled *)
	bAxis10Coupled				:BOOL;					(* Axis coupled *)
END_VAR
VAR
	(* Enummerations *)

	(* Variables *)

	(* References *)

	(* Interfaces *)

	(* Instances *)

END_VAR


IF NOT bEnable							(* Signal FB enable *)
THEN
	F_ChkAllAxisCoupled := FALSE;

	RETURN;
END_IF

F_ChkAllAxisCoupled := bAxis1Coupled
					   AND bAxis2Coupled
					   AND bAxis3Coupled
					   AND bAxis4Coupled
					   AND bAxis5Coupled
					   AND bAxis6Coupled
					   AND bAxis7Coupled
					   AND bAxis8Coupled
					   AND bAxis9Coupled
					   AND bAxis10Coupled;

END_FUNCTION

// ---- POUs/Tc3 Objects/Automation/Axis/F_ChkAllAxisEnabled_1.TcPOU
FUNCTION F_ChkAllAxisEnabled_1 : BOOL
(*

The function used to detect if all axis controller enabled.

Constructor: 		Patryk Panylo
Company:		E. Riexinger GmbH
Date:			23.04.2015
Version:			1.00

Date:			Revision:		Who:				Comment
dd.mm.yyyy		x.xx			Initials			comment

*)
VAR_INPUT
	(* Input variables / Eingang Variablen *)
	bEnable						:BOOL;						(* Signal FB enable *)
	bEnabledAxis1				:BOOL;						(* Controller enabled *)
	bEnabledAxis2				:BOOL;						(* Controller enabled *)
	bEnabledAxis3				:BOOL;						(* Controller enabled *)
	bEnabledAxis4				:BOOL;						(* Controller enabled *)
	bEnabledAxis5				:BOOL;						(* Controller enabled *)
	bEnabledAxis6				:BOOL;						(* Controller enabled *)
	bEnabledAxis7				:BOOL;						(* Controller enabled *)
	bEnabledAxis8				:BOOL;						(* Controller enabled *)
	bEnabledAxis9				:BOOL;						(* Controller enabled *)
	bEnabledAxis10				:BOOL;						(* Controller enabled *)
END_VAR
VAR
	(* Enummerations *)

	(* Variables *)

	(* References *)

	(* Interfaces *)

	(* Instances *)

END_VAR


IF NOT bEnable							(* Signal FB enable *)
THEN
	F_ChkAllAxisEnabled := FALSE;

	RETURN;
END_IF

F_ChkAllAxisEnabled := bEnabledAxis1
					  AND bEnabledAxis2
					  AND bEnabledAxis3
					  AND bEnabledAxis4
					  AND bEnabledAxis5
					  AND bEnabledAxis6
					  AND bEnabledAxis7
					  AND bEnabledAxis8
					  AND bEnabledAxis9
					  AND bEnabledAxis10;

END_FUNCTION

// ---- POUs/Tc3 Objects/Automation/Axis/F_ChkAllAxisInSamePos_1.TcPOU
FUNCTION F_ChkAllAxisInSamePos_1 : BOOL
(*

The function used to detect if all axis have the same position.

Constructor: 		Patryk Panylo
Company:		E. Riexinger GmbH
Date:			09.07.2016
Version:			1.00

Date:			Revision:		Who:				Comment
dd.mm.yyyy		x.xx			Initials			comment

*)
VAR_INPUT
	(* Input variables / Eingang Variablen *)
	bEnable						:BOOL;					(* Signal FB enable *)
	lrAxis1Pos					:LREAL;					(* Axis position [mm] *)
	lrAxis2Pos					:LREAL;					(* Axis position [mm] *)
	lrAxis3Pos					:LREAL;					(* Axis position [mm] *)
	lrAxis4Pos					:LREAL;					(* Axis position [mm] *)
	lrAxis5Pos					:LREAL;					(* Axis position [mm] *)
	lrAxis6Pos					:LREAL;					(* Axis position [mm] *)
	lrAxis7Pos					:LREAL;					(* Axis position [mm] *)
	lrAxis8Pos					:LREAL;					(* Axis position [mm] *)
	lrAxis9Pos					:LREAL;					(* Axis position [mm] *)
	lrAxis10Pos					:LREAL;					(* Axis position [mm] *)
	lrTolerance					:LREAL := 2;					(* Tolerance [mm] *)
END_VAR
VAR
	(* Enummerations *)

	(* Variables *)
	nIdx1						:INT;
	nIdx2						:INT;
	arlrAxisPos					:ARRAY[1..10] OF LREAL;

	(* References *)

	(* Interfaces *)

	(* Instances *)

END_VAR


IF NOT bEnable							(* Signal FB enable *)
THEN
	F_ChkAllAxisInSamePos := TRUE;

	RETURN;
END_IF

arlrAxisPos[1] := lrAxis1Pos;
arlrAxisPos[2] := lrAxis2Pos;
arlrAxisPos[3] := lrAxis3Pos;
arlrAxisPos[4] := lrAxis4Pos;
arlrAxisPos[5] := lrAxis5Pos;
arlrAxisPos[6] := lrAxis6Pos;
arlrAxisPos[7] := lrAxis7Pos;
arlrAxisPos[8] := lrAxis8Pos;
arlrAxisPos[9] := lrAxis9Pos;
arlrAxisPos[10] := lrAxis10Pos;

F_ChkAllAxisInSamePos := TRUE;

FOR nIdx1 := 1 TO 10 DO
	FOR nIdx2 := 1 TO 10 DO
		IF ABS(arlrAxisPos[nIdx1] - arlrAxisPos[nIdx2]) > lrTolerance
		THEN
			F_ChkAllAxisInSamePos := FALSE;
			EXIT;
		END_IF
	END_FOR
END_FOR;

END_FUNCTION

// ---- POUs/Tc3 Objects/Automation/Axis/F_ChkAllAxisNotMoving_1.TcPOU
FUNCTION F_ChkAllAxisNotMoving_1 : BOOL
(*

The function used to detect if all axis not moving.

Constructor: 		Patryk Panylo
Company:		E. Riexinger GmbH
Date:			23.04.2015
Version:			1.00

Date:			Revision:		Who:				Comment
dd.mm.yyyy		x.xx			Initials			comment

*)
VAR_INPUT
	(* Input variables / Eingang Variablen *)
	bEnable						:BOOL;						(* Signal FB enable *)
	bAxis1NotMoving				:BOOL;						(* Axis not moving *)
	bAxis2NotMoving				:BOOL;						(* Axis not moving *)
	bAxis3NotMoving				:BOOL;						(* Axis not moving *)
	bAxis4NotMoving				:BOOL;						(* Axis not moving *)
	bAxis5NotMoving				:BOOL;						(* Axis not moving *)
	bAxis6NotMoving				:BOOL;						(* Axis not moving *)
	bAxis7NotMoving				:BOOL;						(* Axis not moving *)
	bAxis8NotMoving				:BOOL;						(* Axis not moving *)
	bAxis9NotMoving				:BOOL;						(* Axis not moving *)
	bAxis10NotMoving			:BOOL;						(* Axis not moving *)
END_VAR
VAR
	(* Enummerations *)

	(* Variables *)

	(* References *)

	(* Interfaces *)

	(* Instances *)

END_VAR


IF NOT bEnable							(* Signal FB enable *)
THEN
	F_ChkAllAxisNotMoving := FALSE;

	RETURN;
END_IF

F_ChkAllAxisNotMoving := bAxis1NotMoving
					   AND bAxis2NotMoving
					   AND bAxis3NotMoving
					   AND bAxis4NotMoving
					   AND bAxis5NotMoving
					   AND bAxis6NotMoving
					   AND bAxis7NotMoving
					   AND bAxis8NotMoving
					   AND bAxis9NotMoving
					   AND bAxis10NotMoving;

END_FUNCTION

// ---- POUs/Tc3 Objects/Automation/Axis/F_ChkAllAxisReferenced_1.TcPOU
FUNCTION F_ChkAllAxisReferenced_1 : BOOL
(*

The function used to detect if all axis referenced.

Constructor: 		Patryk Panylo
Company:		E. Riexinger GmbH
Date:			23.04.2015
Version:			1.00

Date:			Revision:		Who:				Comment
dd.mm.yyyy		x.xx			Initials			comment

*)
VAR_INPUT
	(* Input variables / Eingang Variablen *)
	bEnable						:BOOL;						(* Signal FB enable *)
	bReferencedAxis1				:BOOL;						(* Controller referenced *)
	bReferencedAxis2				:BOOL;						(* Controller referenced *)
	bReferencedAxis3				:BOOL;						(* Controller referenced *)
	bReferencedAxis4				:BOOL;						(* Controller referenced *)
	bReferencedAxis5				:BOOL;						(* Controller referenced *)
	bReferencedAxis6				:BOOL;						(* Controller referenced *)
	bReferencedAxis7				:BOOL;						(* Controller referenced *)
	bReferencedAxis8				:BOOL;						(* Controller referenced *)
	bReferencedAxis9				:BOOL;						(* Controller referenced *)
	bReferencedAxis10			:BOOL;						(* Controller referenced *)
END_VAR
VAR
	(* Enummerations *)

	(* Variables *)

	(* References *)

	(* Interfaces *)

	(* Instances *)

END_VAR


IF NOT bEnable                          (* Signal FB enable *)
THEN
	F_ChkAllAxisReferenced := FALSE;

	RETURN;
END_IF;

F_ChkAllAxisReferenced := bReferencedAxis1
						AND bReferencedAxis2
						AND bReferencedAxis3
						AND bReferencedAxis4
						AND bReferencedAxis5
						AND bReferencedAxis6
						AND bReferencedAxis7
						AND bReferencedAxis8
						AND bReferencedAxis9
						AND bReferencedAxis10;

END_FUNCTION

// ---- POUs/Tc3 Objects/Automation/Axis/F_ChkAllAxisStandStill_1.TcPOU
FUNCTION F_ChkAllAxisStandStill_1 : BOOL
(*

The function used to detect if all axis stand still.

Constructor: 		Patryk Panylo
Company:		E. Riexinger GmbH
Date:			23.04.2015
Version:			1.00

Date:			Revision:		Who:				Comment
dd.mm.yyyy		x.xx			Initials			comment

*)
VAR_INPUT
	(* Input variables / Eingang Variablen *)
	bEnable						:BOOL;					(* Signal FB enable *)
	bAxis1StandStill				:BOOL;					(* Axis stand still *)
	bAxis2StandStill				:BOOL;					(* Axis stand still *)
	bAxis3StandStill				:BOOL;					(* Axis stand still *)
	bAxis4StandStill				:BOOL;					(* Axis stand still *)
	bAxis5StandStill				:BOOL;					(* Axis stand still *)
	bAxis6StandStill				:BOOL;					(* Axis stand still *)
	bAxis7StandStill				:BOOL;					(* Axis stand still *)
	bAxis8StandStill				:BOOL;					(* Axis stand still *)
	bAxis9StandStill				:BOOL;					(* Axis stand still *)
	bAxis10StandStill				:BOOL;					(* Axis stand still *)
END_VAR
VAR
	(* Enummerations *)

	(* Variables *)

	(* References *)

	(* Interfaces *)

	(* Instances *)

END_VAR


IF NOT bEnable							(* Signal FB enable *)
THEN
	F_ChkAllAxisStandStill := FALSE;

	RETURN;
END_IF

F_ChkAllAxisStandStill := bAxis1StandStill
					   AND bAxis2StandStill
					   AND bAxis3StandStill
					   AND bAxis4StandStill
					   AND bAxis5StandStill
					   AND bAxis6StandStill
					   AND bAxis7StandStill
					   AND bAxis8StandStill
					   AND bAxis9StandStill
					   AND bAxis10StandStill;

END_FUNCTION

// ---- POUs/Tc3 Objects/Automation/Axis/F_ChkAxisError.TcPOU
FUNCTION F_ChkAxisError : BOOL
(*

The function used to detect if any error existss.

Constructor: 		Patryk Panylo
Company:		E. Riexinger GmbH
Date:			23.04.2015
Version:			1.00

Date:			Revision:		Who:				Comment
dd.mm.yyyy		x.xx			Initials			comment

*)
VAR_INPUT
	(* Input variables / Eingang Variablen *)
	bEnable						:BOOL;						(* Signal FB enable *)
	bAxis1Error					:BOOL;						(* Axis error *)
	bAxis2Error					:BOOL;						(* Axis error *)
	bAxis3Error					:BOOL;						(* Axis error *)
	bAxis4Error					:BOOL;						(* Axis error *)
	bAxis5Error					:BOOL;						(* Axis error *)
	bAxis6Error					:BOOL;						(* Axis error *)
	bAxis7Error					:BOOL;						(* Axis error *)
	bAxis8Error					:BOOL;						(* Axis error *)
	bAxis9Error					:BOOL;						(* Axis error *)
	bAxis10Error				:BOOL;						(* Axis error *)
END_VAR
VAR
	(* Enummerations *)

	(* Variables *)

	(* References *)

	(* Interfaces *)

	(* Instances *)

END_VAR


IF NOT bEnable							(* Signal FB enable *)
THEN
	F_ChkAxisError := bEnable;

	RETURN;
END_IF

F_ChkAxisError := bAxis1Error
				  OR bAxis2Error
				  OR bAxis3Error
				  OR bAxis4Error
				  OR bAxis5Error
				  OR bAxis6Error
				  OR bAxis7Error
				  OR bAxis8Error
				  OR bAxis9Error
				  OR bAxis10Error;

END_FUNCTION

// ---- POUs/Tc3 Objects/Automation/Cylinder/FB_Cylinder_1.TcPOU
FUNCTION_BLOCK FB_Cylinder_1
(*
Base class of cylinder.
Cylinder control two directions with handshake.

Constructor: 		Patryk Panylo
Company:		E. Riexinger GmbH
Date:			06.03.2013
Version:			1.00

Date:			Revision:		Who:				Comment
10.30.2013		.02				PPA					Error diagnose off
10.02.2015		.03				PPA					Move in manual in spite of error
13.05.2016		.04				PPA					Valve Off if came limit imput, Control outputs dependent on input state
10.09.2019		.05				PPA					Safety
10.06.2020		.05				PPA					In first cycle check inf move to base or move to work
*)
VAR_INPUT
	(* Input variables / Eingang Variablen *)
	bEnable						:BOOL;			(* Signal FB enable *)
	bAirPressure				:BOOL;			(* Signal air pressure *)
	bSafetyOk					:BOOL;			(* Safety OK  *)
	bReset						:BOOL;			(* Signal reset *)
	bAutoHand					:BOOL;			(* Auto := TRUE, Hand := FALSE *)
	bHandBase					:BOOL;			(* Move hand to base position *)
	bHandWork					:BOOL;			(* Move hand to work position *)
	bAutoBase					:BOOL;			(* Move auto to base position *)
	bAutoWork					:BOOL;			(* Move auto to work position *)
	bBasePos					:BOOL;			(* Base position *)
	bWorkPos					:BOOL;			(* Work position *)
	bAtBasePos					:BOOL;			(* At base position *)
	bAtWorkPos					:BOOL;			(* At work position *)
	bBaseRelease				:BOOL;			(* Base position release *)
	bWorkRelease				:BOOL;			(* Work position release *)
	bControlStateOn				:BOOL;			(* TRUE - control with input state *)
	bControlOff					:BOOL;			(* TRUE - controle off *)
	bValveOff					:BOOL;			(* TRUE -  valve off with limit input *)
	bValveErrOff				:BOOL;			(* TRUE -  valve off if error *)
	bErrorOff					:BOOL;			(* TRUE - error diagnose off *)
	tTimeOut					:TIME := T#5s;	(* TimeOut *)
END_VAR
VAR_OUTPUT
	(* Output variables / Ausgang Variablen *)
	bMoveToBase					:BOOL;			(* Move to base position *)
  	bMoveToWork					:BOOL;			(* Move to work position *)
	bEndBase					:BOOL;			(* Base position reached *)
  	bEndWork					:BOOL;			(* Work position reached *)
 	bNoEndPos					:BOOL;			(* End position not reached *)
	bSafetyLock					:BOOL;			(* Lock safety because of moving *)
	bError						:BOOL;			(* Error *)
	udnErrorNo					:UDINT;			(* Error number *)
	sErrorMsg					:STRING; 		(* Error message *)
END_VAR
VAR_IN_OUT
	(* Input Output variables / Ausgang Variablen *)
	bHomeCompleted				:BOOL;			(* Home completed *)
END_VAR
VAR
	(* Enummerations *)

	(* Variables *)
	bFirstBase					:BOOL;
	bFirstWork					:BOOL;
	bTargetBase					:BOOL;
	bTargetWork					:BOOL;

	bFirstTime					:BOOL;
	(* References *)

	(* Interfaces *)

	(* Instances *)
	rtHandBase					:R_TRIG;
	rtHandWork					:R_TRIG;
	rtAutoBase					:R_TRIG;
	rtAutoWork					:R_TRIG;

	tonFirstTime				:TON;		
 	tonWatchDog					:TON;
END_VAR

IF NOT bEnable
THEN
	bMoveToBase := FALSE;			(* Move to base position *)
  	bMoveToWork := FALSE;			(* Move to work position *)
	bEndBase := FALSE;				(* Base position reached *)
  	bEndWork := FALSE;				(* Work position reached *)
	bError := FALSE;
	udnErrorNo := 0;					(* Error number *)
	sErrorMsg := ''; 					(* Error message *)
	tonWatchDog(IN := FALSE);
	bFirstTime := FALSE;
	RETURN;
END_IF


IF NOT bFirstTime
THEN
	bMoveToBase := FALSE;			(* Move to base position *)
  	bMoveToWork := FALSE;			(* Move to work position *)
	bFirstBase := bBasePos AND NOT bWorkPos;
	bFirstWork := NOT bBasePos AND bWorkPos;
	bTargetBase := FALSE;
	bTargetWork := FALSE;
	bEndBase := FALSE;				(* Base position reached *)
  	bEndWork := FALSE;				(* Work position reached *)
	bFirstTime := TRUE;
	RETURN;
END_IF;

(* Air pressure ok / Luftdruck ok *)
IF NOT bAirPressure
THEN
	rtHandBase(CLK:= FALSE);
	rtHandWork(CLK:= FALSE);
	bSafetyLock := FALSE;
	RETURN;
END_IF;

(* Safety lock *)
bSafetyLock := bHandBase
			  OR bHandWork;

A_SetInputs();
A_ChkOpMode();
A_SetOutputs();
A_Status();

ACTION A_ChkOpMode:

(* Check operating mode *)
IF bAutoHand					(* Automatic *)
THEN
	IF rtAutoBase.Q
	     AND NOT bError
	THEN
		bTargetBase := TRUE;
		bTargetWork := FALSE;
	END_IF;

	IF rtAutoWork.Q
 	     AND NOT bError
	THEN
		bTargetBase := FALSE;
		bTargetWork := TRUE;
	END_IF;

ELSE						(* Manual *)
	IF rtHandBase.Q
	    AND bBaseRelease
	    (* AND NOT bError *)
	THEN
		bTargetBase := TRUE;
		bTargetWork := FALSE;
	END_IF;

	IF rtHandWork.Q
	    AND bWorkRelease
	    (* AND NOT bError *)
	THEN
		bTargetBase := FALSE;
		bTargetWork := TRUE;
	END_IF

END_IF;

tonFirstTime(
	IN := bTargetBase AND bTargetWork,	  
	PT := T#2S
);

IF tonFirstTime.Q
THEN
	IF bFirstBase
	THEN
		bTargetBase := FALSE;
		bFirstBase := FALSE;
	ELSIF bFirstWork
	THEN
		bTargetWork := FALSE;
		bFirstWork := FALSE;
	END_IF	
END_IF
END_ACTION

ACTION A_SetInputs:

(* Check inputs  *)
rtHandBase(CLK:= bHandBase AND bSafetyOk);
rtHandWork(CLK:= bHandWork AND bSafetyOk);
rtAutoBase(CLK:= bAutoBase AND bBaseRelease AND bSafetyOk);
rtAutoWork(CLK:= bAutoWork AND bWorkRelease AND bSafetyOk);
END_ACTION

ACTION A_SetOutputs:

(* Set outputs move to base position  *)
IF bBaseRelease
     OR bAtBasePos
THEN
	IF  bTargetBase
	     AND NOT bMoveToBase
	THEN
		bMoveToBase := TRUE;
		bMoveToWork := FALSE;
		tonWatchDog(IN := FALSE);
	END_IF;

ELSE
	IF bTargetBase
	     AND  bMoveToBase
	THEN
		bMoveToBase := FALSE;

		IF NOT bAutoHand
		THEN
			bTargetBase := FALSE;
		END_IF;

	END_IF;
END_IF;

(* Set outputs move to work position  *)
IF bWorkRelease
    OR bAtWorkPos
THEN
	IF  bTargetWork
	     AND NOT bMoveToWork
	THEN
		bMoveToBase := FALSE;
		bMoveToWork := TRUE;
		tonWatchDog(IN := FALSE);
	END_IF;

ELSE
	IF bTargetWork
	     AND  bMoveToWork
	THEN
		bMoveToWork := FALSE;

		IF NOT bAutoHand
		THEN
			bTargetWork := FALSE;
		END_IF;

	END_IF;
END_IF;

IF NOT bAutoHand
    AND (bMoveToBase
         OR bMoveToWork)
THEN
	bHomeCompleted := FALSE;
END_IF;
END_ACTION

ACTION A_Status:

(* Error reset *)
IF bReset
     AND bError
THEN
	udnErrorNo := 0;					(* Error number *)
	sErrorMsg := ''; 					(* Error message *)
	tonWatchDog(IN := FALSE);
END_IF;

(* Timer starts when cylinder is not  in base and work position *)
tonWatchDog(IN := NOT bErrorOff
				 AND (
					(bMoveToWork AND NOT bAtWorkPos)
				   	OR (bMoveToBase AND NOT bAtBasePos)
				   	OR (NOT bAtBasePos AND NOT bAtWorkPos)
				   	OR (bAtBasePos AND bAtWorkPos)),
			PT := tTimeOut);

(* Error if cylinder does not reach base or work position*)
IF tonWatchDog.Q 
   AND NOT bError
THEN
	IF bMoveToWork
	THEN
		IF NOT bAtWorkPos AND NOT bAtBasePos
		THEN
			udnErrorNo := 1; 								(* Set error number *)
			sErrorMsg := 'Work position not reached';
		ELSIF NOT bAtWorkPos AND bAtBasePos
		THEN
			udnErrorNo := 2; 								(* Set error number *)
			sErrorMsg := 'Not move in work position';
		ELSIF bAtWorkPos AND bAtBasePos
		THEN
			udnErrorNo := 5; 									(* Set error number *)
			sErrorMsg := 'Both position reached';
		END_IF
	ELSIF bMoveToBase
	THEN
		IF NOT bAtWorkPos AND NOT bAtBasePos
		THEN
			udnErrorNo := 3; 								(* Set error number *)
			sErrorMsg := 'Base position not reached';
		ELSIF bAtWorkPos AND NOT bAtBasePos
		THEN
			udnErrorNo := 4; 								(* Set error number *)
			sErrorMsg := 'Not move in base position';
		ELSIF bAtWorkPos AND bAtBasePos
		THEN
			udnErrorNo := 5; 									(* Set error number *)
			sErrorMsg := 'Both position reached';
		END_IF
	ELSIF bAtWorkPos AND bAtBasePos
	THEN
		udnErrorNo := 5; 									(* Set error number *)
		sErrorMsg := 'Both position reached';
	END_IF
END_IF

bError := udnErrorNo <> 0;


(* End base position reached  *)
bEndBase := bAtBasePos
		        AND NOT bAtWorkPos
		        AND NOT bError;

(* End wrok position reached  *)
bEndWork := NOT bAtBasePos
		        AND bAtWorkPos
		        AND NOT bError;

(* End position not reached *)
IF bTargetBase
THEN
	bNoEndPos := NOT bAtBasePos;

ELSIF bTargetWork
THEN
	bNoEndPos :=  NOT bAtWorkPos;

ELSE
	bNoEndPos := FALSE;
END_IF


(* Valve off if error  *)
IF bError
     AND (bMoveToBase OR bMoveToWork)
     AND bValveErrOff
THEN
	bMoveToBase := FALSE;
	bMoveToWork := FALSE;
	bTargetBase := FALSE;
	bTargetWork := FALSE;
END_IF;

(* Control with input state *)
IF bControlStateOn
THEN
	IF bAutoHand					(* Automatic *)
	THEN
		IF NOT bAutoBase
		THEN
			bMoveToBase := FALSE;
			bTargetBase := FALSE;
		END_IF

		IF NOT bAutoWork
		THEN
			bMoveToWork := FALSE;
			bTargetWork := FALSE;
		END_IF
	
	ELSE						(* Manual *)
		IF NOT bHandBase
		THEN
			bMoveToBase := FALSE;
			bTargetBase := FALSE;
		END_IF

		IF NOT bHandWork
		THEN
			bMoveToWork := FALSE;
			bTargetWork := FALSE;
		END_IF
	
	END_IF;
END_IF

(* Check control off *)
IF bControlOff
    AND (
		bMoveToBase OR bMoveToWork
		OR bTargetBase OR bTargetWork
	      )
THEN
	bMoveToBase := FALSE;
	bMoveToWork := FALSE;
	bTargetBase := FALSE;
	bTargetWork := FALSE;
END_IF

(* Check valve off *)
IF bValveOff
THEN
	IF bAtBasePos
	    AND (bMoveToBase OR bTargetBase)
	THEN
		bMoveToBase := FALSE;
		bTargetBase := FALSE;

	ELSIF bAtWorkPos
	    	   AND (bMoveToWork OR bTargetWork)
	THEN
		bMoveToWork := FALSE;
		bTargetWork := FALSE;
	END_IF
END_IF
END_ACTION

END_FUNCTION_BLOCK

// ---- POUs/Tc3 Objects/Automation/Force/FB_ForceController_1.TcPOU
FUNCTION_BLOCK FB_ForceController_1
(*

The function block used to 

Constructor: 		Patryk Panylo
Company:		E. Riexinger GmbH
Date:			17.02.2016
Version:			1.00

Date:			Revision:		Who:				Comment

*)
VAR_INPUT
	(* Input variables / Eingang Variablen *)
	bEnable					:BOOL;					(* Signal FB enable *)
	bControllerOn				:BOOL;					(* Controler on *)
	lrVeloKp					:LREAL := 0.1;				(* Kp Proportionalfaktor, deltaF x Kp -> v *)
	lrVeloTi					:LREAL := 10000;			(* Ti Integrationsfaktor*)
	lrPreCtrlVelo				:LREAL := 0.01;			(* Feedforward velocity precontrol wieghting =  0..1 *)
	lrPVForce				:LREAL;					(* Process variable of force *)
	lrSPForce				:LREAL;					(* Set point of force *)
	lrMaxForce				:LREAL;					(* Maximum force *)
	lrDeltaMax				:LREAL := 0.01;
	lrVeloMax				:LREAL := 10.0;			(* Maximum velocity [%] *)
	lrVeloMin				:LREAL := 0.0;				(* Minimum velocity [%] *)
	lrTaskCycle				:LREAL;					(* Task cycle *)
END_VAR
VAR_OUTPUT
	(* Output variables / Ausgang Variablen *)
	lrCVVelo					:LREAL;					(* Controller value of velocity [%] *)
END_VAR
VAR_IN_OUT
	(* Input Output variables / Ausgang Variablen *)

END_VAR
VAR
	(* Enummerations *)

	(* Variables *)

	(* References *)

	(* Interfaces *)

	(* Instances *)
	fbActForceFilter				:FB_ValueFilter;					(* Actual position filter *)
	fbCtrlPID						:FB_CtrlPID;

END_VAR
VAR CONSTANT

END_VAR


IF NOT bEnable
THEN
	lrCVVelo := 100;
	RETURN;
END_IF

(* Current force value filtering *)
fbActForceFilter(
	bEnable := TRUE,
	lrInSignal := lrPVForce,
	lrDeltaMax := lrDeltaMax,
);

IF bControllerOn
     AND fbActForceFilter.lrOutSignal < lrMaxForce
THEN

	fbCtrlPID(
		bEnable := TRUE,
		lrSetPoint := lrSPForce,
		lrProcessVariable := fbActForceFilter.lrOutSignal,
		lrDeadZone := 1.0,
		lrSignalOffset := 0.0,
		lrKp := lrVeloKp,
		lrTi := lrVeloTi,
		lrTd := 0.0,
		lrTaskCycle := lrTaskCycle,
		bManual := ,
		lrManualSignal:= ,
		lrLimitMin := lrVeloMin,
		lrLimitMax := lrVeloMax,
		lrProcessErr => ,
		bLimitMin => ,
		bLimitMax => );

	(*lrCVVelo := MAX(0.0, (fbCtrlPID.lrCtrlVariable * (1.0 - MIN(lrPreCtrlVelo, 1))) + (fbActForceFilter.lrOutSignal * MIN(lrPreCtrlVelo, 1))); (* where lrPreCtrlVelo := 0.01 *)*)
	lrCVVelo := MAX(0.0, (fbCtrlPID.lrCtrlVariable * (1.0 - MIN(lrPreCtrlVelo, 1))) + (lrCVVelo * MIN(lrPreCtrlVelo, 1)));				       (* where lrPreCtrlVelo := 0.99 *)

ELSE
	lrCVVelo := 0.0;
END_IF

END_FUNCTION_BLOCK

// ---- POUs/Tc3 Objects/Automation/Force/FB_ForceReg_1.TcPOU
FUNCTION_BLOCK FB_ForceReg_1
VAR_INPUT
	rVelocityMax			:REAL := 10.0;
	rVelocityMin			:REAL := 0.0;
	PID_Reg: FB_PID_Regler;
	SollForceInt: INT := 20;
	IstForceInt: INT := 20;
	bRegelung: BOOL := FALSE;
	PWM_Aus: INT := 0;
	Force_Aus: REAL := 0.0;
	Simulation: BOOL := FALSE;
END_VAR
VAR_OUTPUT
	ForceOK: BOOL := FALSE;
	ForceOn: BOOL := FALSE;
	ForceLeistung: REAL := 0.0;
END_VAR
VAR
	PWM_Inc: INT := 0;
	PWM_Max: INT := 200;
	ForceModellReal: REAL := 0.0;
	K_Modell: REAL := 0.1;
	K_Modell_EM: REAL := 0.9;
	Force_Normal: REAL := 19.0;
	ForceModellInt: INT := 0;
	T_Modell: REAL := 360.0;
	bfirstCycle: BOOL := TRUE;
END_VAR

IF bFirstCycle THEN 				 (* Anfangsinitialisierungen *)

	PWM_Inc := 0;

	PID_Reg	(	
		fMax:=INT_TO_REAL(PWM_Max) ,
		fMin := 0.0,
		fD_Max := 1.0E10,
		fD_Min := -1.0E10,
		fKr := 1.0,
		fTN := 0.0,
		fTv := 0.0,
		fTau := 0.0,
		fOff := 0.0,
		fTab := 2.0,
		fState :=0.0,
		fIntegral := 0.0,
		fSoll := 0.0,
		fIst := 0.0
	);

	K_Modell 		:= EXP(-0.01/T_Modell);
	K_Modell_EM 	:= 1.0 - K_Modell;
	
	bFirstCycle:=FALSE;
END_IF

(* Zähler füR PID 0 incrementieren *)
PWM_Inc := 	PWM_Inc  + 1;

(* Regelung für PID 0 aufrufen *)
IF (PWM_Inc >= PWM_Max ) 
THEN
	PWM_Inc :=  0;

	(* Hier Regler einbauen *)
	IF bRegelung 
	THEN
		IF Simulation 
		THEN
			PID_Reg(fSoll:=SollForceInt, fIst:=ForceModellInt);
		ELSE
			PID_Reg(fSoll:=SollForceInt, fIst:=IstForceInt);
		END_IF
	
		PWM_Aus :=  REAL_TO_INT(PID_Reg.fAus);
		Force_Aus :=  PID_Reg.fAus;
		ForceOK := PID_Reg.bRegOK;
	ELSE
		PID_Reg.fIntegral := 0.0;
		PID_Reg(fSoll:=0.0, fIst:=0.0);
		PWM_Aus :=  0;
		Force_Aus :=  0.0;
		ForceOK := TRUE;
	
	END_IF

	IF ( PWM_Aus > PWM_Max ) THEN PWM_Aus:= PWM_Max; END_IF
	IF ( PWM_Aus < 0      ) THEN PWM_Aus := 0; END_IF

	IF ( Force_Aus > rVelocityMax ) THEN Force_Aus := rVelocityMax; END_IF
	IF ( Force_Aus < rVelocityMin ) THEN Force_Aus := rVelocityMin; END_IF

END_IF

(* PWM für PID  ausgeben == Inaktivierungsstrecke*)

ForceOn := FALSE;
IF (  PWM_Aus > PWM_Inc ) 
THEN		
	ForceOn := TRUE;        
END_IF

IF Simulation
THEN
	ForceModellReal := K_Modell*ForceModellReal;
	IF (  PWM_Aus > PWM_Inc ) THEN		ForceModellReal := K_Modell_EM*ForceModellReal;       END_IF
	ForceModellReal  := ForceModellReal + Force_Normal;
	ForceModellInt	:=REAL_TO_INT(ForceModellReal*10.0);
END_IF

END_FUNCTION_BLOCK

// ---- POUs/Tc3 Objects/Automation/Force/FB_PID_Regler_1.TcPOU
FUNCTION_BLOCK FB_PID_Regler_1
VAR_INPUT
	fSoll: REAL;
	fIst: REAL;
	fMax: REAL := 1.0;
	fMin: REAL := 0.0;
	fD_Max: REAL := 1.0;
	fD_Min: REAL := 0.0;
	fKr: REAL;
	fTn: REAL;
	fTv: REAL;
	fTau: REAL;
	fOff: REAL;
	fTab: REAL;
	fState: REAL;
	fIntegral: REAL;
END_VAR
VAR_OUTPUT
	bRegOK: BOOL := FALSE;
	fAus: REAL;
END_VAR
VAR
	fU: REAL;
	fU_Max: REAL;
	fU_Min: REAL;
	fU_Pd: ARRAY[1..2] OF REAL;
	fU_I: ARRAY[1..2] OF REAL;
	fE: ARRAY[1..4] OF REAL;
	fP: ARRAY[1..2] OF REAL;
	fQ: ARRAY[1..6] OF REAL;
	cMax: REAL;
	cMin: REAL;
	cD_Max: REAL := 1.0;
	cD_Min: REAL := 0.0;
	cKr: REAL;
	cTn: REAL;
	cTv: REAL;
	cTau: REAL;
	cOff: REAL;
	cTab: REAL;
	cState: REAL;
	cIntegral: REAL;
	nReg_Typ: INT;
	RegMaxAbweichung: REAL := 20.0;
END_VAR
VAR CONSTANT
	D_REG_I :INT:= 0;
	D_REG_M :INT := 1;
	D_REG_V :INT := 2;
	D_REG :INT := 4;
	I_REG :INT:= 8;
	P_REG :INT := 16;
	PD_I_REG :INT := 20;
	PD_M_REG :INT := 21;
	PD_V_REG :INT := 22;
	PI_REG :INT := 24;
	PID_I_REG :INT := 28;
	PID_M_REG :INT := 29;
	PID_V_REG :INT := 30;
	SET_MIN_MAX :INT := 101;
	ReglerResetState :INT := 102;
	ReglerInit :INT := 103;
	ReglerSet :INT := 104;
	ReglerCalculate :INT := 105;
END_VAR


IF (cMax  <>  fMax) 	THEN cMax := fMax; 	END_IF		 (*  Maximum                            *)
IF (cMin  <>  fMin) 	THEN cMin := fMin; 	END_IF	 	 (*  Minimum                            *)
IF (cD_Max  <>  fD_Max) 	THEN cD_Max := fD_Max; 	END_IF	 	 (*  Maximum der Änderung               *)
IF (cD_Min  <>  fD_Min) 		THEN cD_Min := fD_Min; 	END_IF	 	  (*  Minimum der Änderung               *)

IF ( (cState <>  fState) OR (cIntegral <>  fIntegral)) 		THEN
	cState := fState;
	cIntegral := fIntegral;
	fU := cState;
	fU_I[1] := fU_I[2] := cIntegral;
	fU_Pd[2] := fU_Pd[1] := 0.0;
	fE[4]		:=	fE[3]	:=	fE[2]		:=	fE[1]		:= 	0.0;
END_IF	 	  (*   Änderung Integral      *)

IF (  (cKr  <>  fKr) OR (cTn <> fTn) OR (cTv <> fTv) OR (cTau <> fTau)  OR (cOff <> fOff) OR (cTab <> fTab) ) THEN

     		cKr  := fKr;      (*  Verstärkung                       *)
		cTn  := fTn;      (*  Nachstellzeit                     *)
    		cTv  := fTv;      (*  Vorstellzeit                      *)
    		cTau := fTau;    (*  Tau                               *)
    		cOff := fOff;     (*  Offset                            *)

    		cTab := fTab;

(*    ReglerResetState(0.0, 0.0, p_r);           (*** Rücksetzen der Reglergrößen ***) *)
                  IF ( cTn = 0.0 ) THEN 	fU := fU_I[1] := fU_I[2] := 	fU_Pd[2] := fU_Pd[1] := 	fE[4]		:=	fE[3]	:=	fE[2]		:=	fE[1]		:= 	0.0;  END_IF

    		fP[1] := fP[2] := 0;         (*** Rücksetzen der Parameter ***)
    		fQ[1] := fQ[2] := fQ[3] := fQ[4] := fQ[5] := fQ[6] := 0;

    		nReg_Typ := 0;
    		IF ( cKr > 0 ) THEN nReg_Typ := nReg_Typ + P_REG;   END_IF  (*** Ermittlung der Reglertyps***)
    		IF ( cTn > 0 ) THEN nReg_Typ := nReg_Typ +  I_REG; END_IF
    		IF ( cTv > 0 ) THEN
      			 nReg_Typ := nReg_Typ + D_REG;
       			IF (cTau = 0) THEN nReg_Typ := nReg_Typ + D_REG_I;  END_IF(*** Ideale Differenz ***)
       			IF (cTau <  0) THEN nReg_Typ := nReg_Typ + D_REG_M;  END_IF(*** Gemittelte Differenz ***)
       			IF (cTau >  0) THEN nReg_Typ := nReg_Typ + D_REG_V;  END_IF(*** Verzögerte Differenz ***)
    		END_IF

		CASE nReg_Typ OF                  (*** Berechnung der Parameter ***)
		    P_REG :        (*** P-Regler ***********************************)
		       fQ[1] := cKr;
		    PI_REG :       (*** PI-Regler **********************************)
		       fQ[1] := cKr;

		       fQ[6] := cKr*cTab/cTn;
		    PD_I_REG :     (*** PD-Regler,      ideale Differenz  **********)
		       fQ[1] :=  cKr*cTv/cTab + cKr;
		       fQ[2] := -cKr*cTv/cTab;
		    PD_M_REG :     (*** PD-Regler,  gemittelte Differenz  **********)
		       fQ[1] :=  cKr*(1.0+cTv/6.0/cTab);
		       fQ[2] :=  cKr*cTv/2.0/cTab;
		       fQ[3] := -fQ[2];
		       fQ[4] :=  fQ[3]/3;
		    PD_V_REG :     (*** PD-Regler,  verzögerte Differenz  **********)
		       fP[1] := EXP(-cTab/cTau);

		       fQ[1] :=   cKr + cKr*cTv/cTau;
		       fQ[2] :=  -cKr - cKr*cTv/cTau + cKr*(1.0 - fP[1]) ;
		    PID_I_REG :    (*** PID-Regler,     ideale Differenz  **********)
		       fQ[1] :=  cKr*cTv/cTab + cKr;
		       fQ[2] := -cKr*cTv/cTab;

		       fQ[6] :=  cKr*cTab/cTn;
		    PID_M_REG :    (*** PID-Regler, gemittelte Differenz  **********)
		       fQ[1] :=  cKr*cTv/6/cTab + cKr;
		       fQ[2] :=  cKr*cTv/2/cTab;
		       fQ[3] := -fQ[2];
		       fQ[4] :=  fQ[3]/3;

		       fQ[6] :=  cKr*cTab/cTn;
		    PID_V_REG :    (*** PID-Regler, verzögerte Differenz  **********)
		       fP[1] :=  EXP(-cTab/cTau);

		       fQ[1] :=   cKr + cKr*cTv/cTau;
		       fQ[2] :=  -cKr - cKr*cTv/cTau + cKr*(1.0 - fP[1]) ;

		       fQ[6] :=  cKr*cTab/cTn;
		    I_REG :        (*** I-Regler ***********************************)
		       fQ[6] :=  cTab/cTn;

		END_CASE
END_IF


	fE[1] := fSoll - fIst;       	   (*** Regelabweichung ***)
	IF ( ABS(fE[1]) < RegMaxAbweichung ) THEN bRegOK := TRUE; ELSE bRegOK := FALSE; END_IF

	fU_Max := fU + cD_Max;   (*** dynamische Stellbegrenzung ***)
	IF (fU_Max > cMax) THEN fU_Max := cMax; END_IF

    	fU_Min := fU + cD_Min;
	IF (fU_Min < cMIN) THEN fU_Min := cMIN; END_IF
			                                          (*** Reglergleichung füR P- und D-Anteil***)
    	fU := fU_Pd[1] := fP[1]*fU_Pd[2] +   fQ[1]*fE[1] + fQ[2]*fE[2] +  fQ[3]*fE[3] + fQ[4]*fE[4];

                                          (*** Reglergleichung mit altem I-Anteil***)
    	fU := fU + fU_I[2];
                                      (*** Begrenzung der Stellgröße ***)
    	IF ( fU  > (fU_Max - cOff) ) THEN
             fU := fU_Max - cOff;
	ELSE
         		IF ( fU < (fU_Min - cOff) ) THEN
                		fU := fU_Min - cOff;
	         ELSE
                                          (*** Reglergleichung für I-Anteil***)
			fU_I[1] := fU_I[2] + fQ[6]*fE[1];
                                          (*** Gesamt-Reglergleichung ***)
			fU := (fU_Pd[1] + fU_I[1]);

                                      (*** Begrenzung der Stellgröße ***)
			IF ( fU > (fU_Max - cOff) ) THEN
                   		fU := fU_Max - cOff;
	                   	fU_I[1]  := fU - fU_Pd[1];
			ELSE
         		          	IF ( fU < (fU_Min - cOff) ) THEN
                   			fU := fU_Min - cOff;
		         		         fU_I[1]  := fU - fU_Pd[1];
	         		      	END_IF
         		   	END_IF
         		END_IF
    	END_IF                                          (*** Umspeichern der Regelgrößen ***)
	fU_Pd[2] := fU_Pd[1];
	fU_I[2]  := fU_i[1];

	fE[4] := fE[3];
	fE[3] := fE[2];
	fE[2] := fE[1];

                                        (*** Übergabe der Stellgröße ***)
	fAus := fU + cOff;

END_FUNCTION_BLOCK

// ---- POUs/Tc3 Objects/Automation/OperationMode/FB_ModeSelector_1.TcPOU
FUNCTION_BLOCK FB_ModeSelector_1
(*

The function block used to control opration mode.

Constructor: 		Patryk Panylo
Company:		E. Riexinger GmbH
Date:			23.04.2015
Version:			1.00

Date:			Revision:		Who:				Comment
dd.mm.yyyy		x.xx			Initials			comment

*)
VAR_INPUT
	(* Input variables / Eingang Variablen *)
	bStart					:BOOL;						(* Signal start *)
	bStop					:BOOL;						(* Signal stop *)
	bAbort					:BOOL;						(* Signal abort *)
	bHome					:BOOL;						(* Signal home *)
	bReference				:BOOL;						(* Signal reference *)
	bReset					:BOOL;						(* Signal reset *)
	bAutoStartRelease		:BOOL;						(* Auto start release *)
	bHomeStartRelease		:BOOL;						(* Home start release *)
	bMaintenanceStartRelease:BOOL;						(* Maintenance start release *)
	bAutoToHome				:BOOL;						(* If auto completed go to home *)
	bChangeModeWithHome		:BOOL;						(* If mode was changed start home *)
	bHomeCompleted			:BOOL;						(* Home completed *)
	bAutoCompleted			:BOOL;						(* Auto completed *)
	bMaintenanceCompleted	:BOOL;						(* Maintenance completed *)
	bAllDoorsClosed 		:BOOL;						(* All doors closed *)
	bAllDoorsLocked 		:BOOL;						(* All doors locked *)
	bLightCurtainOk			:BOOL;						(* Light curtain ok *)
END_VAR
VAR_OUTPUT
	(* Output variables / Ausgang Variablen *)
	etMachineMode			:ET_MachineMode;			(* Machine mode enum variable *)
	etMachineState			:ET_MachineState;			(* Machine state enum variable *)
	etMaintenanceType		:ET_MaintenanceType;		(* Maintenance type enum variable *)
	bModeAutomatic			:BOOL;						(* Machine mode automatic *)
	bModeHome				:BOOL;						(* Machine mode home *)
	bModeManual				:BOOL;						(* Machine mode manual *)
	bModeMaintenance		:BOOL;						(* Machine mode maintenance *)
	bMachineRunning			:BOOL;						(* Machine running *)
	bMachineStandstill		:BOOL;						(* Machine standstill *)
	bConfirmAlarm			:BOOL;						(* Confirm alarm *)
END_VAR
VAR_IN_OUT
	etMachineModeReq		:ET_MachineMode;			(* Machine mode request enum variable *)
	etMaintenanceTypeReq	:ET_MaintenanceType;		(* Maintenance type request *)
END_VAR
VAR
	(* Enummerations *)

	(* Variables *)
	etMachinePrvState		:ET_MachineState;			(* Machine previous active state enum variable *)
	etMachinePrvModeReq		:ET_MachineMode;			(* Machine mode request previous enum variable *)
	
	bModeExecute			:BOOL;						(* Mode execute *)
	bSafetyCompleted		:BOOL;						(* Safety completed *)
	
	bFirstHomeCompleted		:BOOL;						(* First home is completed *)	
	(* References *)

	(* Interfaces *)

	(* Instances *)
	rtStart					:R_TRIG;
	rtStop					:R_TRIG;
	rtAbort					:R_TRIG;

END_VAR


bConfirmAlarm := bReset;
bSafetyCompleted := bAllDoorsLocked				(* Safety completed *)
				      AND bLightCurtainOk;

etMaintenanceType := etMaintenanceTypeReq;					  
					  
IF bHome
THEN
	etMachineModeReq := ET_MachineMode_eHome;
END_IF;

IF bMaintenanceCompleted
THEN
	etMachineModeReq := ET_MachineMode_eManual;
END_IF

IF bHomeCompleted
THEN
	bFirstHomeCompleted := bHomeCompleted;

	IF etMachineMode = ET_MachineMode_eHome                          	 (* Set auto mode *)
	    AND etMachinePrvState <> ET_MachineState_eAutoExe
	    AND etMachinePrvState <> ET_MachineState_eAutoSteppingExe
	    AND etMachinePrvState <> ET_MachineState_eAutoSteppingNoExe
		AND etMachinePrvState <> ET_MachineState_eMaintenanceExe
	    AND bModeExecute
	THEN
		IF etMachinePrvModeReq = ET_MachineMode_eManual
		THEN
			etMachineModeReq := ET_MachineMode_eManual;
			etMachinePrvModeReq := ET_MachineMode_eUndefined;
		ELSE
			etMachineModeReq := ET_MachineMode_eAutomatic;
		END_IF
	END_IF;	
ELSE
	IF etMachineModeReq <> ET_MachineMode_eManual                   	 (* Set home mode *)
	   AND SEL(bFirstHomeCompleted, TRUE, etMachineModeReq <> ET_MachineMode_eMaintenance)
	THEN
		etMachineModeReq := ET_MachineMode_eHome;
	
	END_IF;
END_IF;

IF (etMachineModeReq <> etMachineMode)                                    		(* Stop always if changed mode *)
THEN
	(*bStart := FALSE *)
	bStop := TRUE;
	
	IF (etMachineMode = ET_MachineMode_eAutomatic
	      AND etMachineModeReq = ET_MachineMode_eStepping)
	     OR
	     (etMachineMode = ET_MachineMode_eStepping
	      AND etMachineModeReq = ET_MachineMode_eAutomatic)
		  OR
	     (etMachineMode = ET_MachineMode_eManual
	      AND etMachineModeReq = ET_MachineMode_eMaintenance)
	THEN
		bStop := FALSE;
		
	ELSIF ((etMachineMode = ET_MachineMode_eAutomatic
			OR etMachineMode = ET_MachineMode_eStepping
			OR etMachineMode = ET_MachineMode_eCycle)
			AND bMachineRunning
			AND bChangeModeWithHome)
	THEN
		bStart := TRUE;
		bStop := FALSE;
		etMachinePrvModeReq := etMachineModeReq;
		etMachineModeReq := ET_MachineMode_eHome;
			
	END_IF;
	
	etMachineMode := etMachineModeReq;

END_IF;

rtStart(CLK := bStart);								(* Check start *)

rtStop(CLK := bStop								(* Check stop *)
		        OR bAbort
		        OR bAutoCompleted
		        OR (NOT bSafetyCompleted AND bMachineRunning));
rtAbort(CLK := bAbort);

IF rtStop.Q
THEN
	bModeExecute := FALSE;

	IF bAutoToHome
	     AND bAutoCompleted
	THEN
		etMachineModeReq := ET_MachineMode_eHome;
	END_IF
	
	IF etMachinePrvModeReq = ET_MachineMode_eManual
		OR etMachineMode = ET_MachineMode_eMaintenance
	THEN
		etMachineModeReq := ET_MachineMode_eManual;
		etMachinePrvModeReq := ET_MachineMode_eUndefined;
	END_IF

ELSIF rtStart.Q
	    AND bAllDoorsClosed
	    AND bLightCurtainOk
	    AND NOT bStop
	    AND NOT bAbort
	    AND ((etMachineMode = ET_MachineMode_eMaintenance 
			  AND SEL(etMachineState = ET_MachineState_eMaintenanceExe, 
					  bMaintenanceStartRelease, TRUE))
	    	  OR (etMachineMode = ET_MachineMode_eHome 
			  AND SEL(etMachineState = ET_MachineState_eHomeExe 
					  OR etMachineState = ET_MachineState_eHomeRefExe, 
					  bHomeStartRelease, TRUE))
	    	  OR ((etMachineMode = ET_MachineMode_eAutomatic OR etMachineMode = ET_MachineMode_eStepping) 
				   AND SEL(etMachineState = ET_MachineState_eAutoExe 
						   OR etMachineState = ET_MachineState_eAutoSteppingExe 
						   OR etMachineState = ET_MachineState_eAutoSteppingNoExe,
						   bAutoStartRelease, TRUE)))
THEN
	bModeExecute := TRUE;

END_IF;

bStart := FALSE;
bStop := FALSE;

CASE etMachineMode
OF
	ET_MachineMode_eAutomatic:            (* Statement section automatic *)
		bModeAutomatic := TRUE;
		bModeHome := FALSE;
		bModeManual := FALSE;
		bModeMaintenance := FALSE;

		IF bModeExecute
		     AND bSafetyCompleted
		THEN
			etMachineState := ET_MachineState_eAutoExe;
			etMachinePrvState := etMachineState;
		ELSE
		 	etMachineState := ET_MachineState_eIdle;
		END_IF;
	    
	ET_MachineMode_eStepping:             (* Statement section stepping *)
		bModeAutomatic := TRUE;
		bModeHome := FALSE;
		bModeManual := FALSE;
		bModeMaintenance := FALSE;

		IF bModeExecute
		     AND bSafetyCompleted
		THEN
			IF rtStart.Q
			THEN
				etMachineState := ET_MachineState_eAutoSteppingExe;
			ELSE
				etMachineState := ET_MachineState_eAutoSteppingNoExe;
			END_IF;

			etMachinePrvState := etMachineState;
		ELSE
			etMachineState := ET_MachineState_eIdle;
		END_IF;

	ET_MachineMode_eHome:                 (* Statement section home  *)
		bModeAutomatic := FALSE;
		bModeHome := TRUE;
		bModeManual := FALSE;
		bModeMaintenance := FALSE;
		
		IF bModeExecute
		     AND bSafetyCompleted
		THEN
			IF bReference
			THEN
				etMachineState := ET_MachineState_eHomeRefExe;
			ELSE
				etMachineState := ET_MachineState_eHomeExe;
			END_IF;

			etMachinePrvState := etMachineState;
		ELSE
			etMachineState := ET_MachineState_eIdle;
		END_IF;

	ET_MachineMode_eManual:              (* Statement section manual  *)
		bModeExecute := FALSE;
		bModeAutomatic := FALSE;
		bModeHome := FALSE;
		bModeManual := TRUE;
		bModeMaintenance := FALSE;

		etMachineState := ET_MachineState_eIdle;

	ET_MachineMode_eMaintenance:              (* Statement section maintenance  *)
		bModeAutomatic := FALSE;
		bModeHome := FALSE;
		bModeManual := FALSE;
		bModeMaintenance := TRUE;
	
		IF bModeExecute
		     AND bSafetyCompleted
		THEN
			etMachineState := ET_MachineState_eMaintenanceExe;
			etMachinePrvState := etMachineState;
		ELSE
		 	etMachineState := ET_MachineState_eIdle;
		END_IF;
	
	ELSE
		bModeExecute := FALSE;
		bModeAutomatic := FALSE;
		bModeHome := FALSE;
		bModeManual := FALSE;
		bModeMaintenance := FALSE;
	    
	    etMachineState := ET_MachineState_eUndefined;
        
END_CASE;

bMachineRunning := bModeExecute
		           AND etMachineMode <> ET_MachineMode_eManual
		           AND etMachineMode <> ET_MachineMode_eIdle
		           AND etMachineMode <> ET_MachineMode_eUndefined;
                    
bMachineStandstill := NOT bMachineRunning;

END_FUNCTION_BLOCK

// ---- POUs/Tc3 Objects/Automation/Override/FB_OverrideSelection_1.TcPOU
FUNCTION_BLOCK FB_OverrideSelection_1
(*

The function block used to select override of axis.

Constructor: 		Patryk Panylo
Company:		E. Riexinger GmbH
Date:			23.04.2015
Version:			1.00

Date:			Revision:		Who:				Comment
dd.mm.yyyy		x.xx			Initials			comment

*)
VAR_INPUT
	(* Input variables / Eingang Variablen *)
	bEnable						:BOOL;						(* Signal FB enable *)
	rGlobalOverride				:REAL;						(* Global override *)
	rAcc							:REAL;						(* Accerlation of Override [%/s] *)
	rDec						:REAL;						(* Decerlation of Override [%/s] *)
END_VAR
VAR_OUTPUT
	(* Output variables / Ausgang Variablen *)
	rActOverride					:REAL;						(* Actual override *)
	bActGlobalOverride			:BOOL;						(* Actual override is global *)
	bActLocalOverride			:BOOL;						(* Actual override is local *)
END_VAR
VAR_IN_OUT
	(* Input Output variables / Ausgang Variablen *)
	rLocalOverride				:REAL;						(* Actual override *)
END_VAR
VAR
	(* Enummerations *)

	(* Variables *)
	rCacheGlobalOverride			:REAL;						(* Caches global override *)
	rCacheLocalOverride			:REAL;						(* Caches local override *)

	bFirstTime					:BOOL;						(* First run *)

	(* References *)

	(* Interfaces *)

	(* Instances *)
	tonChkCycleTime				:TON;						(* Check cycle time *)
END_VAR
VAR CONSTANT

END_VAR


IF NOT bEnable
THEN
	bFirstTime := FALSE;                               		(* Firstrun *)
	rActOverride := 0.0;                               		(* Override to set *)
	bActGlobalOverride := FALSE;                       	(* Actual override is global *)
	bActLocalOverride := FALSE;                       	(* Actual override is local *)
	RETURN;
END_IF;

IF NOT bFirstTime
THEN
	rCacheGlobalOverride := rGlobalOverride;          	(* Cache values *)
	rCacheLocalOverride := rLocalOverride;            		(* Cache values *)
	bActGlobalOverride := TRUE;                        			(* Actual override is global *)
	bActLocalOverride := FALSE;                       			(* Actual override is local *)
	bFirstTime := TRUE;                                				(* Firstrun *)
END_IF;

A_SelectLocal();
A_SelectGlobal();

ACTION A_SelectGlobal:

IF rCacheGlobalOverride <> rGlobalOverride
    OR rLocalOverride >= rGlobalOverride
THEN
	rCacheGlobalOverride := rGlobalOverride;
	rActOverride := rGlobalOverride;
	bActGlobalOverride := TRUE;                       	 		(* Actual override is global *)
	bActLocalOverride := FALSE;                        			(* Actual override is local *)
	rLocalOverride := rGlobalOverride;                		(* Set local Override *)
	rCacheLocalOverride := rGlobalOverride;           		(* Set local Override *)
END_IF;
END_ACTION

ACTION A_SelectLocal:

IF rCacheLocalOverride <> rLocalOverride
    AND rLocalOverride < rGlobalOverride
THEN
	rCacheLocalOverride := rLocalOverride;
	rActOverride := rLocalOverride;
	bActGlobalOverride := FALSE;                       			(* Actual override is global *)
	bActLocalOverride := TRUE;                        			(* Actual override is local *)
END_IF;
END_ACTION

END_FUNCTION_BLOCK

// ---- POUs/Tc3 Objects/Automation/Override/FB_Override_1.TcPOU
FUNCTION_BLOCK FB_Override_1
(*

The function block used to control override of axis.

Constructor: 		Patryk Panylo
Company:		E. Riexinger GmbH
Date:			23.04.2015
Version:			1.00

Date:			Revision:		Who:				Comment
dd.mm.yyyy		x.xx			Initials			comment

*)
VAR_INPUT
	(* Input variables / Eingang Variablen *)
	bEnable						:BOOL;						(* Signal FB enable *)
	bBypassAccDec				:BOOL;						(* Bypassing acceleratin und deceleration rActOverride = rSetOverride *)
	bSetOverideMax				:BOOL;						(* Set maximum override *)
	rAcc							:REAL;						(* Accerlation of Override [%/s] *)
	rDec						:REAL;						(* Decerlation of Override [%/s] *)
END_VAR
VAR_OUTPUT
	(* Output variables / Ausgang Variablen *)
	rActOverride					:REAL;						(* Actual Override *)
END_VAR
VAR_IN_OUT
	rSetOverride					:REAL;						(* Set Override *)
END_VAR
VAR
	(* Enummerations *)

	(* Variables *)
	rSetOverrideInternal			:REAL;						(* Internal Set Override limited *)
	rAccOverridePerCycle			:REAL;						(* Override accerleration per cycle *)
	rDecOverridePerCycle			:REAL;						(* Override deceleration per cycle *)
	tCycleTime					:TIME;						(* Detected cycle Time *)
	bFirstTime					:BOOL;						(* First run *)

	(* References *)

	(* Interfaces *)

	(* Instances *)
	tonChkCycleTime				:TON;						(* Check cycle time *)
	rtSetOverideMax				:R_TRIG;
END_VAR
VAR CONSTANT
	rMIN_OVERRIDE				:REAL := 0.0;					(* Minimum override *)
	rMAX_OVERRIDE				:REAL := 100.0;				(* Maximum override *)
	rACC_MIN					:REAL := 0.1;					(* Minimum accerleration *)
	rDEC_MIN					:REAL := 0.1;					(* Minimum decerleration *)
	tMAX_CYCLE_TIME			:TIME := t#1s;					(* Maximum cycle time *)
END_VAR

IF NOT bEnable
THEN
	bFirstTime := FALSE;								(* First run *)
	rActOverride := 100.0;								(* Set Override *)
	RETURN;
END_IF;

IF NOT bFirstTime                                             					 (* First run after bEnable *)
THEN
	tonChkCycleTime(					   				 (* Start Timer to check  cycle time *)
		IN := TRUE,
		PT := tMAX_CYCLE_TIME
	);
	
	IF tonChkCycleTime.ET <> t#0s                              			 (* Timer was running one circle *)
	THEN
		tCycleTime := tonChkCycleTime.ET;                     		 (* Detectet circle time *)

		tonChkCycleTime(					 			 (* Stop Timer *)
			IN := FALSE,
			PT := tMAX_CYCLE_TIME
		);

		bFirstTime := TRUE;                                     			(* First run *)
	END_IF;
END_IF;

(* Set max overide *)
rtSetOverideMax(CLK := bSetOverideMax);
IF rtSetOverideMax.Q
THEN
	rSetOverride := rMAX_OVERRIDE;
END_IF

(* Check Limits *)
rSetOverrideInternal := LIMIT(                      					 (* Internal Override Limited *)
	rMIN_OVERRIDE,              							 (* Minimum Override *)
	rSetOverride,              							 	 (* Set Override *)
	rMAX_OVERRIDE               							 (* Maximum Overide *)
);

IF bBypassAccDec
THEN
	rActOverride := rSetOverrideInternal;                  			 (* Actual Override = Set Override *)
ELSE
	IF tCycleTime <> t#0s
	THEN

		A_Acceleration();

		A_Deceleration();

	END_IF;
END_IF;

ACTION A_Acceleration:

IF rSetOverrideInternal > rActOverride                          	(* Override has to be added *)
THEN
	(* Check if accerlaeration zero *)
	IF rAcc <= 0
	THEN
		rAcc := rACC_MIN;                                         	(* Set accerlaeration to minimum *)
	END_IF;

	(* Calculate Accerleration per cycle *)
	rAccOverridePerCycle := rAcc / (TIME_TO_REAL(tMAX_CYCLE_TIME)
							     / TIME_TO_REAL(tCycleTime));
	
	rActOverride := rActOverride + rAccOverridePerCycle;        (* Add Override *)
	IF rActOverride > rSetOverrideInternal                      		 (* Actoverride  run over Set Override ? *)
	THEN
		rActOverride := rSetOverrideInternal;             (* Set  Override equal *)
	END_IF;
END_IF;
END_ACTION

ACTION A_Deceleration:

IF rSetOverrideInternal < rActOverride                             (* Override has to subed *)
THEN
	(* Check if decerlaeration zero *)
	IF rDec <= 0
	THEN
		rDec := rDEC_MIN;                                         	(* Set decerlaeration to minimum *)
	END_IF;

	(* Calculate decerleration per cycle *)
	rDecOverridePerCycle := rDec / (TIME_TO_REAL(tMAX_CYCLE_TIME) /
								TIME_TO_REAL(tCycleTime));
	
	rActOverride := rActOverride - rDecOverridePerCycle;        (* Sub Override *)
	IF rActOverride < rSetOverrideInternal                        		 (* Actoverride  run over Set Override ? *)
	THEN
	    rActOverride := rSetOverrideInternal;                  (* Set  Override equal *)
	END_IF;
END_IF;
END_ACTION

END_FUNCTION_BLOCK

// ---- POUs/Tc3 Objects/Automation/Process/FB_StartProcess_1.TcPOU
FUNCTION_BLOCK FB_StartProcess_1
(*

The function block used to control start process.

Constructor: 		Patryk Panylo
Company:		E. Riexinger GmbH
Date:			27.04.2015
Version:			1.00

Date:			Revision:		Who:				Comment
dd.mm.yyyy		x.xx			Initials			comment

*)
VAR_INPUT
	(* Input variables / Eingang Variablen *)
	bEnable						:BOOL;						(* Enable FB signal *)
	bStart						:BOOL;						(* Signal start *)
	bStop						:BOOL;						(* Signal stop *)
	bDone						:BOOL;						(* Signal done *)
	bStepping					:BOOL;						(* Stepping active *)
END_VAR
VAR_OUTPUT
	(* Output variables / Ausgang Variablen *)
	bStartProcess				:BOOL;						(* Start process *)
END_VAR
VAR_IN_OUT
	(* Input Output variables / Ausgang Variablen *)
	bHomeCompleted				:BOOL;			(* Home completed *)
END_VAR
VAR
	(* Enummerations *)

	(* Variables *)

	(* References *)

	(* Interfaces *)

	(* Instances *)
	rtStart						:R_TRIG;
END_VAR

IF NOT bEnable
THEN
	rtStart(CLK := FALSE);
	bStartProcess := FALSE;
	RETURN;
END_IF;


(* Start process with handshake *)
rtStart(CLK:= bStart);

IF (bDone
    OR bStop
    OR NOT bHomeCompleted)
    AND bStartProcess
THEN
	bStartProcess := FALSE;

ELSIF rtStart.Q
      AND NOT bStartProcess
THEN
	IF bStepping
	THEN
		 bStartProcess := rtStart.Q;
	ELSE
		bStartProcess := TRUE;
	END_IF;
END_IF;

END_FUNCTION_BLOCK

// ---- POUs/Tc3 Objects/Automation/Spindle/FB_CoolingDevice_1.TcPOU
FUNCTION_BLOCK FB_CoolingDevice_1
(*

The function block used to control power supply.

Constructor: 		Patryk Panylo
Company:		E. Riexinger GmbH
Date:			23.04.2015
Version:			1.00

Date:			Revision:		Who:				Comment
dd.mm.yyyy		x.xx			Initials			comment

*)
VAR_INPUT
	(* Input variables / Eingang Variablen *)
	bEnable					:BOOL;						(* Enable FB signal *)
	bIn						:BOOL;						(* Input signal *)
	tCoolingDeviceOn			:TIME := t#2s;					(* Timeout power supply on *)
	tCoolingDeviceOff			:TIME := t#1s;					(* Timeout power supply off *)
END_VAR
VAR_OUTPUT
	(* Output variables / Ausgang Variablen *)
	bOut					:BOOL;						(* Air pressure ok *)
	bError					:BOOL;						(* Error by no air pressure *)
	udnErrorNo				:UDINT;
	udnMessageNo			:UDINT;
	sMsg					:STRING;
END_VAR
VAR_IN_OUT

END_VAR
VAR
	(* Enummerations *)

	(* Variables *)
	bFirstTime				:BOOL;						(* First cycle *)

	(* References *)

	(* Interfaces *)

	(* Instances *)
	tonCoolingDeviceOn		:TON;						(* Timer to delay *)
	tofCoolingDeviceOff		:TOF;						(* Timer to delay *)
	tCoolingDevice			:BOOL;
END_VAR

IF NOT bEnable
THEN
	bOut := TRUE;
	bError := FALSE;
	udnErrorNo := 0;
	udnMessageNo := 0;
	sMsg := '';
	tonCoolingDeviceOn(IN := FALSE,
				            PT := tCoolingDeviceOn);
	tofCoolingDeviceOff(IN := FALSE,
	            			 PT := tCoolingDeviceOff);
	bFirstTime := FALSE;
    RETURN;
END_IF;

IF NOT bFirstTime
THEN
	bError := FALSE;
	udnErrorNo := 0;
	udnMessageNo := 0;
	sMsg := '';
	tonCoolingDeviceOn(IN := FALSE,
	          			  PT := tCoolingDeviceOn);
	tofCoolingDeviceOff(IN := FALSE,
	             			 PT := tCoolingDeviceOff);
	bFirstTime := TRUE;
END_IF;

(* Timer starts when came rising edge of signal *)
tonCoolingDeviceOn(
	IN := bIn,
         PT := tCoolingDeviceOn
);

tofCoolingDeviceOff(
	IN := bIn,
         PT := tCoolingDeviceOff
);

bOut := tonCoolingDeviceOn.Q;
bError := NOT tofCoolingDeviceOff.Q;

IF bError
THEN
	udnErrorNo := 1;
	udnMessageNo := 0;
	sMsg := 'No power supply';
ELSE
	udnErrorNo := 0;
	udnMessageNo := 0;
	sMsg := '';
END_IF;

END_FUNCTION_BLOCK

// ---- POUs/Tc3 Objects/Automation/Vacuum/FB_Vacuum_1.TcPOU
FUNCTION_BLOCK FB_Vacuum_1
(*
Base class of vacuum.

Constructor: 		Patryk Panylo
Company:		E. Riexinger GmbH
Date:			13.05.2016
Version:			1.01

Date:			Revision:		Who:				Comment
27.10.2016		.01				PPA					Monitoring of pump engine


*)
VAR_INPUT
	(* Input variables / Eingang Variablen *)
	bEnable						:BOOL;			(* Signal FB enable *)
	bAirPressure				:BOOL;			(*  Signal air pressure *)
	bSafetyOk					:BOOL;			(* Safety OK  *)
	bEngineOk					:BOOL;			(*  Pump engine is ok *)
	bReset						:BOOL;			(*  Signal reset *)
	bAutoHand 					:BOOL;			(*  Auto := TRUE, Hand := FALSE *)
	bHandOpen					:BOOL;			(*  Hand open *)
	bHandClose					:BOOL;			(*  Hand close *)
	bAutoOpen					:BOOL;			(*  Auto open *)
	bAutoClose					:BOOL;			(*  Auto close *)
	bOpened						:BOOL;			(* Valve opened *)
	bClosed						:BOOL;			(* Valve closed *)
	bOpenRelease 				:BOOL;			(* Open release *)
	bCloseRelease				:BOOL;			(* Close release *)
	bControlStateOn				:BOOL;			(* TRUE - control with input state *)
	bControlOff					:BOOL;			(* TRUE - controle off *)
	tControlOff					:TIME;			(* Time > 0 delay to control off *)
	bValveErrOff				:BOOL;			(* TRUE -  valve off if error *)
	bErrorOff					:BOOL;			(* TRUE - error diagnose off *)
	tTimeOut					:TIME := T#5S;	(* TimeOut *)
END_VAR
VAR_OUTPUT
	(* Output variables / Ausgang Variablen *)
	bOpen						:BOOL;			(* Valve open *)
	bClose						:BOOL;			(* Valve close *)
	bEndOpened					:BOOL;			(* Open reached *)
	bEndClosed					:BOOL;			(* Close reached *)
	bNoEndPos					:BOOL;			(* End position not reached *)
	bSafetyLock					:BOOL;			(* Lock safety because of moving *)
	bError						:BOOL;			(* Error *)
	udnErrorNo					:UDINT;			(* Error number *)
	sErrorMsg					:STRING;		(* Error message *)
END_VAR
VAR_IN_OUT
	(* Input Output variables / Ausgang Variablen *)
	bHomeCompleted				:BOOL;			(* Home completed *)
END_VAR
VAR
	tonWatchDog					:TON;
	rtHandOpen					:R_TRIG;
	rtHandClose					:R_TRIG;
	rtAutoOpen					:R_TRIG;
	rtAutoClose					:R_TRIG;
	tonControlOff					:TON;
	bTargetOpen					:BOOL;
	bTargetClose					:BOOL;
	bFirstTime					:BOOL;

END_VAR


IF NOT bEnable
THEN
	bOpen := FALSE;                  		(* Valve open *)
	bClose := FALSE;				(* Valve close *)
	bEndOpened := FALSE;               	(* Valve opended *)
	bEndClosed := FALSE;               	(* Valve closed *)
	bError := FALSE;
	udnErrorNo := 0;                   		(* Error number *)
	sErrorMsg := '';                   		(* Error message *)

	tonWatchDog(
		IN := FALSE,
	         PT := tTimeOut
	);
	tonControlOff(
		IN := FALSE,
	         PT := tControlOff
	);

	bFirstTime := FALSE;
	RETURN;
END_IF;


IF NOT bFirstTime
THEN
	bOpen := FALSE;                    		(* Valve open *)
	bClose := FALSE;                  		(* Valve close *)
	bEndOpened := FALSE;              	(* Valve opended *)
	bEndClosed := FALSE;               	(* Valve closed *)
	bFirstTime := TRUE;
	RETURN;
END_IF;


(* Air pressure ok / Luftdruck ok *)
IF NOT bAirPressure
     OR NOT bEngineOk
THEN
	bOpen := FALSE;
	bClose := FALSE;
	bTargetOpen := FALSE;
	bTargetClose := FALSE;
	bSafetyLock := FALSE;
	RETURN;
END_IF;

(* Safety lock *)
bSafetyLock := bHandOpen
			   OR bHandClose;

(* Check inputs  *)
rtHandOpen(CLK := bHandOpen AND bSafetyOk);
rtHandClose(CLK := bHandClose AND bSafetyOk);
rtAutoOpen(CLK := bAutoOpen AND bOpenRelease AND (NOT bControlOff OR tControlOff > T#0MS) AND bSafetyOk);
rtAutoClose(CLK := bAutoClose AND bCloseRelease AND (NOT bControlOff OR tControlOff > T#0MS) AND bSafetyOk);


(* Check operating mode *)
IF bAutoHand                    (* Automatic *)
THEN
	IF rtAutoOpen.Q
	    AND NOT bError
	THEN
		bTargetOpen := TRUE;
		bTargetClose := FALSE;
	END_IF;
	
	IF rtAutoClose.Q
	    AND NOT bError
	THEN
		bTargetOpen := FALSE;
		bTargetClose := TRUE;
	END_IF;
    
ELSE                        (* Manual *)
	IF rtHandOpen.Q
	   AND bOpenRelease
	   (* AND NOT #bError *)
	THEN
		bTargetOpen := TRUE;
		bTargetClose := FALSE;
	END_IF;
	
	IF rtHandClose.Q
	    AND bCloseRelease
	    (* AND NOT #bError *)
	THEN
		bTargetOpen := FALSE;
		bTargetClose := TRUE;
	END_IF;
    
END_IF;


(* Set outputs valve open *)
IF bOpenRelease
THEN
	IF bTargetOpen
	     AND NOT bOpen
	THEN
		bOpen := TRUE;
		bClose := FALSE;
		tonWatchDog(
			IN := FALSE,
			PT := tTimeOut
		);

		tonControlOff(
			IN := FALSE,
			PT := tControlOff
		);
	END_IF;
    
ELSE
	IF bTargetOpen
	    AND bOpen
	THEN
		bOpen := FALSE;
	
		IF NOT bAutoHand
		THEN
		    bTargetOpen := FALSE;
		END_IF;
	
	END_IF;
END_IF;

(* Set outputs valve close *)
IF bCloseRelease
THEN
	IF bTargetClose
	    AND NOT bClose
	THEN
		bOpen := FALSE;
		bClose := TRUE;
		tonWatchDog(
			IN := FALSE,
			PT := tTimeOut
		);

		tonControlOff(
			IN := FALSE,
			PT := tControlOff
		);
	END_IF;
    
ELSE
	IF bTargetClose
	     AND bClose
	THEN
		bClose := FALSE;

		IF NOT bAutoHand
		THEN
			bTargetClose := FALSE;
		END_IF;
	
	END_IF;
END_IF;

IF NOT bAutoHand
     AND (bOpen OR bClose)
THEN
	bHomeCompleted := FALSE;
END_IF;

(* Error reset *)
IF bReset
    AND bError
THEN
	udnErrorNo := 0;                    (* Error number *)
	sErrorMsg := '';                    (* Error message *)
	tonWatchDog(
		IN := FALSE,
	         PT := tTimeOut
	);

END_IF;

(* Timer starts when valve is not opened and work position *)
tonWatchDog(
	IN := NOT bErrorOff
		AND (
			(bClose AND NOT bClosed)
			  OR (bOpen AND NOT bOpened)
			  OR (NOT bOpened AND NOT bClosed)
			  OR (bOpened AND bClosed)),
	PT := tTimeOut
);

(* Error if valve does not reach open or work sensor *)
IF tonWatchDog.Q
    AND NOT bError
THEN
	IF bClose
	THEN
		IF NOT bClosed AND NOT bOpened
		THEN
			udnErrorNo := 1;                                (* Set error number *)
			sErrorMsg := 'Work position not reached';
		ELSIF NOT bClosed AND bOpened
		THEN
			udnErrorNo := 2;                                (* Set error number *)
			sErrorMsg := 'Not move in work position';
		ELSIF bClosed AND bOpened
		THEN
			udnErrorNo := 5;                                    (* Set error number *)
			sErrorMsg := 'Both position reached';
		END_IF;
	ELSIF bOpen
	THEN
		IF NOT bClosed AND NOT bOpened
		THEN
			udnErrorNo := 3;                                (* Set error number *)
			sErrorMsg := 'Base position not reached';
		ELSIF bClosed AND NOT bOpened
		THEN
			udnErrorNo := 4;                                (* Set error number *)
			sErrorMsg := 'Not move in base position';
		ELSIF bClosed AND bOpened
		THEN
			udnErrorNo := 5;                                    (* Set error number *)
			sErrorMsg := 'Both position reached';
		END_IF;
	ELSIF bClosed AND bOpened
	THEN
		udnErrorNo := 5;                                    (* Set error number *)
		sErrorMsg := 'Both position reached';
	END_IF;
END_IF;

bError := udnErrorNo <> 0;

(* Open reached  *)
bEndOpened := bOpened
			    AND NOT bClosed
			    AND NOT bError;

(* Close reached  *)
bEndClosed := NOT bOpened
			  AND bClosed
			  AND NOT bError;

(* End position not reached *)
IF bTargetOpen
THEN
	bNoEndPos := NOT bOpened;
    
ELSIF bTargetClose
THEN
	bNoEndPos := NOT bClosed;

ELSE
    bNoEndPos := FALSE;
END_IF;


(* Valve off if error  *)
IF bError
    AND (bOpen OR bClose)
    AND bValveErrOff
THEN
	bOpen := FALSE;
	bClose := FALSE;
END_IF;

(* Control with input state *)
IF bControlStateOn
THEN
	IF bAutoHand					(* Automatic *)
	THEN
		IF NOT bAutoOpen
		THEN
			bOpen := FALSE;
			bTargetOpen := FALSE;
		END_IF

		IF NOT bAutoClose
		THEN
			bClose := FALSE;
			bTargetClose := FALSE;
		END_IF
	
	ELSE						(* Manual *)
		IF NOT bHandOpen
		THEN
			bOpen := FALSE;
			bTargetOpen := FALSE;
		END_IF

		IF NOT bHandClose
		THEN
			bClose := FALSE;
			bTargetClose := FALSE;
		END_IF
	
	END_IF;
END_IF

(* Check control off *)
IF bControlOff
   AND tControlOff > t#0ms
THEN
	tonControlOff(
		IN := bOpen OR bClose
			 OR bTargetOpen OR bTargetClose,
		PT := tControlOff
	);
    
	IF tonControlOff.Q
	THEN
		bOpen := FALSE;
		bClose := FALSE;
		bTargetOpen := FALSE;
		bTargetClose := FALSE;
	END_IF;
    
ELSE
	tonControlOff(
		IN := FALSE,
		PT := tControlOff
	);
	
	IF bControlOff
	     AND (bOpen OR bClose
		       OR bTargetOpen OR bTargetClose)
	THEN
		bOpen := FALSE;
		bClose := FALSE;
		bTargetOpen := FALSE;
		bTargetClose := FALSE;
	END_IF;
END_IF;

END_FUNCTION_BLOCK

// ---- POUs/Tc3 Objects/Basics/CheckBounds_1.TcPOU
FUNCTION CheckBounds_1 : DINT
VAR_INPUT
	index: DINT;
	lower: DINT;
	upper: DINT;
END_VAR
VAR_EXTERNAL
	fbCheckArrayBounds: FB_CheckArrayBounds;
END_VAR

(*This function checks if an index out of range an array is being accessed *)

fbCheckArrayBounds(
	diArrayIndex			:= index,
	diLowerBound		:= lower,
	diUpperBound		:= upper,
	sLogMessage		=> ,
	diReturnBound		=> CheckBounds);

END_FUNCTION

// ---- POUs/Tc3 Objects/Basics/CheckDivReal_1.TcPOU
FUNCTION CheckDivReal_1 : REAL
VAR_INPUT
	divisor: REAL;
END_VAR
VAR_EXTERNAL
	fbCheckDivRealInfo: FB_CheckDivRealInfo;
END_VAR

(*This function checks if a division by zero is performed*)

fbCheckDivRealInfo(
	rDivisor			:= divisor,
	sLogMessage	=> ,
	rReturnDivReal 	=> CheckDivReal);

END_FUNCTION

// ---- POUs/Tc3 Objects/Basics/FB_CheckArrayBounds_1.TcPOU
FUNCTION_BLOCK FB_CheckArrayBounds_1
VAR_INPUT
	diArrayIndex: DINT;
	diLowerBound: DINT;
	diUpperBound: DINT;
END_VAR
VAR_OUTPUT
	sLogMessage: STRING;
	diReturnBound: DINT;
END_VAR
VAR
	bErrorUpper: BOOL;
	bErrorLower: BOOL;
	fbRTrig_MessageOutputLower: R_TRIG;
	fbRTrig_MessageOutputUpper: R_TRIG;
END_VAR

(*++++++++++ Checkbounds ++++++++++*)
(*If somehow it happens that a value of any of the used arrays that does not exist is being accessed,
the value is either set to the highest declared value (if a value higher than the highest declared value is being accessed) 
or it is set to the lowest declared value (if a value lower than the lowest declared value is being accessed)  *)

IF diArrayIndex< diLowerBound THEN
	diReturnBound:= diLowerBound;
	bErrorLower:= TRUE;

	sLogMessage:= 'CheckBounds: Array index too LOW! Lower Bound: ';			(*Message is put together*)
	sLogMessage:=CONCAT(sLogMessage,DINT_TO_STRING(diLowerBound));
	sLogMessage:=CONCAT(sLogMessage,' Index being accessed: ');
	sLogMessage:=CONCAT(sLogMessage,DINT_TO_STRING(diArrayIndex));

ELSIF diArrayIndex> diUpperBound THEN
	diReturnBound:= diUpperBound;
	bErrorUpper:= TRUE;

	sLogMessage:= 'CheckBounds: Array index too HIGH! Upper Bound: ';			(*Message is put together*)
	sLogMessage:=CONCAT(sLogMessage,DINT_TO_STRING(diUpperBound));
	sLogMessage:=CONCAT(sLogMessage,' Index being accessed: ');
	sLogMessage:=CONCAT(sLogMessage,DINT_TO_STRING(diArrayIndex));

ELSIF NOT (diArrayIndex< diLowerBound) AND
	NOT (diArrayIndex> diUpperBound) THEN
		diReturnBound:= diArrayIndex;
		bErrorUpper:= FALSE;
		bErrorLower:= FALSE;
END_IF

(*++++++++++ ADSLOGDINT ++++++++++*)
(*If somehow it happens that a value of any of the used arrays that does not exist is being accessed,
the Error is written into the Logger Box of the TC System Manager  *)

fbRTrig_MessageOutputLower( CLK:= bErrorLower, Q=> );
fbRTrig_MessageOutputUpper( CLK:= bErrorUpper, Q=> );

IF fbRTrig_MessageOutputLower.Q OR fbRTrig_MessageOutputUpper.Q THEN
	ADSLOGDINT( ADSLOG_MSGTYPE_ERROR OR ADSLOG_MSGTYPE_LOG,sLogMessage,0);	(*Message is written into Event Log*)
END_IF

END_FUNCTION_BLOCK

// ---- POUs/Tc3 Objects/Basics/FB_CheckDivRealInfo_1.TcPOU
FUNCTION_BLOCK FB_CheckDivRealInfo_1
VAR_INPUT
	rDivisor: REAL;
END_VAR
VAR_OUTPUT
	rReturnDivReal: REAL;
	sLogMessage: STRING;
END_VAR
VAR
	bDivisorError: BOOL;
	fbRTrig_MessageOutputDiv: R_TRIG;
END_VAR

IF rDivisor= 0 THEN
	bDivisorError:= TRUE;
	rReturnDivReal:= 1;
ELSE
	rReturnDivReal:= rDivisor;
	bDivisorError:= FALSE;
END_IF

(*++++++++++ ADSLOGDINT ++++++++++*)
(*If somewhere a division by 0 is performed, an Error is written into the Logger Box of the TC System Manager  *)

fbRTrig_MessageOutputDiv( CLK:= bDivisorError, Q=> );

IF fbRTrig_MessageOutputDiv.Q THEN
	sLogMessage:= 'CheckDivReal Error: Division by Zero! Divisor set from 0 to 1. ';					(*Message*)

	ADSLOGDINT( ADSLOG_MSGTYPE_ERROR OR ADSLOG_MSGTYPE_LOG,sLogMessage,0);	(*Message is written into Event Log*)
END_IF

END_FUNCTION_BLOCK

// ---- POUs/Tc3 Objects/Basics/FB_Get_Time_1.TcPOU
FUNCTION_BLOCK FB_Get_Time_1
VAR_INPUT
END_VAR
VAR_OUTPUT
	sDateAndTime: STRING;
END_VAR
VAR
	bBusy: BOOL;
	bError: BOOL;
	udiErrorID: UDINT;
	fbGetTime: NT_GetTime;
	stTime: TIMESTRUCT;
	nStep: UDINT;
	bBlinker: BOOL;
	fbBlinker: FB_Blinker;
	stBlinker:ST_Blinker;
END_VAR

(*This Function Block gets the Windows Systemtime*)

CASE nStep OF
	0:	IF NOT bError AND NOT bBusy THEN
			nStep:= 10;
		ELSE
			nStep:= 30;
		END_IF

	10:	IF stBlinker.Q0 THEN
			fbGetTime.START:= TRUE;
		ELSE
			fbGetTime.START:= FALSE;
			nStep:= 0;
		END_IF

	30:	IF NOT bError AND NOT bBusy THEN
			nStep:= 10;
		END_IF
END_CASE

fbBlinker(tPeriod := t#500ms, stBlinker => stBlinker);

fbGetTime(
			NETID:= '' ,
			START:=   ,
			TMOUT:= DEFAULT_ADS_TIMEOUT ,
			BUSY=> bBusy ,
			ERR=> bError ,
			ERRID=> udiErrorID ,
			TIMESTR=> stTime );

sDateAndTime:= SYSTEMTIME_TO_STRING(stTime);

END_FUNCTION_BLOCK

// ---- POUs/Tc3 Objects/Basics/F_AdsError_Text_1.TcPOU
FUNCTION F_AdsError_Text_1 : STRING
VAR_INPUT
	nCode: UDINT;
END_VAR
VAR
	sText: STRING(255);
END_VAR

